(* IEC 61131-3 sources: daoli-st-library/DL_MathData (part 15) *)

(* ---- FC_DL_HexStringToLword.st ---- *)
(*==============================================================================
 * 组件名称 (Component)  : FC_DL_HexStringToLword
 * 所属子库 (Sublibrary) : DL_MathData
 * 归属目录 (Directory)  : C:\Library\DL_MathData
 * 当前版本 (Version)    : 1.0.0
 * 分类/来源标签         : 函数（FUNCTION）· 纯函数 · 十六进制串解析
 *                         iec-std-wrapper / string / bitstring
 * 兼容性   (Platform)   : CODESYS 3.5 / TwinCAT 3 / 汇川 InoProShop / 施耐德
 *                         Machine Expert；仅用 Standard.library 的 LEN / MID / FIND
 * 溯源声明 (Provenance) : IEC 61131-3 标准语义的道莅防御性实现——内部委托平台标准库语义，
 *                         外围统一错误码 / 钳位 / 双语注释，严禁重实现数学内核。
 * 功能一句话 (Summary)  : 大小写十六进制串解析为 LWORD，奇偶长度、非法字符、
 *                         超长溢出三闸齐备，与 FC_DL_BytesToHexString 互补成对。
 *
 * 功能描述 (Function)   : 一次锁存串长后按序过三闸：长度大于 16 即溢出闸、
 *                         奇数长度即对齐闸、逐字符经三张码表定位失败即非法闸；
 *                         合法路径每字符左移 4 位并入半字节，空串恒等返回零值。
 * 与既有件边界 (Boundary): 本件只解析裸十六进制串，不识别 0x 前缀、不下划线
 *                         分隔；超过 16 个有效位即溢出拒绝，绝不静默截高位。
 * 码位说明 (Codes)      : 信息 16#0002_3040 空输入恒等返回（值零、解析零位）
 *                         故障 16#0002_3041 奇数长度（半个字节无法对齐）
 *                         故障 16#0002_3042 非法字符（不在 0-9 A-F a-f）
 *                         故障 16#0002_3043 超长溢出（有效位大于 16）
 *                         段 16#02_3_40~43 首槽信息级、次槽起故障级。
 * 依赖说明 (Depends)    : 无 DL_ 内部依赖；仅 Standard.library 的 LEN / MID / FIND。
 * 红线自检 (Redline)    : 零全局依赖 ｜ 零 VAR_EXTERNAL ｜ 零 %I/%Q ｜ 纯 IEC 标准库
 *                         移位量 4 恒小于 64 位宽（归一达标）｜ 无除法面
 *                         全变量双语同行注释 ｜ 无定时器实例
 * 修订历史 (Revision)   : 2026-11-18  v1.0.0  首版入库（R32 · 批 1）
 *============================================================================*)

FUNCTION FC_DL_HexStringToLword : BOOL
VAR_INPUT
    sHex : STRING(255);                 // 源十六进制串 [ASCII]，有效位最多 16 / Source hex string, at most 16 digits
END_VAR
VAR_OUTPUT
    uValue  : LWORD;                    // 解析结果 [位串]，域外拒绝时保持零 / Parsed value, zero when refused
    nParsed : INT;                      // 成功解析的有效位数 [位] / Digits parsed on success
    uErrorId: UDINT;                    // 事件码，0 表示无事件 / Event code, zero means none
END_VAR
VAR
    cCh    : STRING(1);   // 当前字符 [字符] / Current character
    nLen   : INT;         // 锁存的源串长度 [字符]，R38 唯一锁存量 / Latched source length
    nVal   : INT;         // 当前半字节值 [值]，域 0 到 15 / Current nibble value, 0 to 15
    nPos   : INT;         // 码表定位结果 [索引]，1 起 / Table position, 1-based
    nI     : INT;         // 字符循环下标 [索引] / Character loop index
    uAcc   : LWORD;       // 累积值 [位串]，出口一次性赋给 uValue / Accumulator
    uCode  : UDINT;       // 码位暂存，出口单点写入 [码] / Code staging
END_VAR
VAR CONSTANT
    DL_HTL_MAXDIG : INT := 16;  // 有效位上限 [位]，LWORD 恰好 64 位 / Digit limit, LWORD is exactly 64 bits
    DL_HTL_ONE    : INT := 1;   // 单字符长度参数 [字符] / Single character length argument
END_VAR

(* 段 1｜输出预置与残留清除 / Pre-set and clear before any branch *)
FC_DL_HexStringToLword := FALSE;
uValue   := 16#0000_0000_0000_0000;
uAcc     := 16#0000_0000_0000_0000;
nParsed  := 0;
uErrorId := 16#0000_0000;
uCode    := 16#0000_0000;

(* 段 2｜LEN 一次锁存 / Latch the length once *)
nLen := LEN(sHex);
IF nLen < 0 THEN
    nLen := 0;                   // 防御：异常返回值钳到零 / Defensive clamp
END_IF

(* 段 3｜空串恒等：信息级告知后成功返回零值 / Empty string identity: inform and succeed *)
IF nLen = 0 THEN
    uErrorId := 16#0002_3040;    // 信息级：空输入恒等返回 / Info: empty input identity
    FC_DL_HexStringToLword := TRUE;
    RETURN;
END_IF

(* 段 4｜溢出闸：有效位超过 16 直接拒绝，绝不静默截高位 / Overflow gate: refuse, never truncate silently *)
IF nLen > DL_HTL_MAXDIG THEN
    uErrorId := 16#0002_3043;    // 故障级：超长溢出 / Fault: overflow by length
    RETURN;
END_IF

(* 段 5｜对齐闸：奇数长度意味着半个字节，解析结果无法定界 / Alignment gate: odd length leaves a half byte undefined *)
IF (nLen MOD 2) = 1 THEN
    uErrorId := 16#0002_3041;    // 故障级：奇数长度 / Fault: odd length
    RETURN;
END_IF

(* 段 6｜逐字符解析：三张码表定位，失败即非法闸 / Parse per character: three tables, failure is the legality gate *)
FOR nI := 1 TO nLen DO
    cCh := MID(sHex, DL_HTL_ONE, nI);                // 取当前字符 / Take the current character
    IF (cCh >= '0') AND (cCh <= '9') THEN
        nPos := FIND('0123456789', cCh);             // 数字表定位，域内恒 1 到 10 / Digit table, 1 to 10
        nVal := nPos - DL_HTL_ONE;                   // 值 0 到 9 / Value 0 to 9
    ELSIF (cCh >= 'A') AND (cCh <= 'F') THEN
        nPos := FIND('ABCDEF', cCh);                 // 大写表定位 / Uppercase table
        nVal := 10 + (nPos - DL_HTL_ONE);            // 值 10 到 15 / Value 10 to 15
    ELSIF (cCh >= 'a') AND (cCh <= 'f') THEN
        nPos := FIND('abcdef', cCh);                 // 小写表定位 / Lowercase table
        nVal := 10 + (nPos - DL_HTL_ONE);            // 值 10 到 15 / Value 10 to 15
    ELSE
        uErrorId := 16#0002_3042;                    // 故障级：非法字符 / Fault: illegal character
        RETURN;
    END_IF
    uAcc := SHL(uAcc, 4) OR INT_TO_LWORD(nVal);      // 左移 4 位并入半字节 / Shift four and OR the nibble
    nParsed := nParsed + DL_HTL_ONE;                 // 有效位计数 / Count the digit
END_FOR

(* 段 7｜出口装配：结果与码位单点写出 / Exit: single write for result and code *)
uValue := uAcc;
uErrorId := uCode;
FC_DL_HexStringToLword := TRUE;
END_FUNCTION

(* ---- FC_DL_HexToStr.st ---- *)
(*
  ==================================================================
  组件名 Component  : FC_DL_HexToStr
  分类   Category   : DL_MathData
  前缀   Naming     : FC_DL_ ｜ b/n/u/f/s/a 类型前缀制（R265）
  版本   Version    : 1.0.0
  功能   Purpose    : 字节串 → HEX 大写文本：每字节展开两位（高半字节
                      在前），输出上限 255 字符（2×127 字节 = 254 字符
                      + $00 终结符），超限按 R49 四步截断样板执行：先判
                      超限并置截断信息码与 bTrunc → 再钳长 → 再写入 →
                      最后显式写 $00 终结符。返回值 = 实际写入字符数
                      （名实双出口）。溯源：本件为「IEC 61131-3 标准语
                      义的道莅防御性实现」，内核委托标准库字符串函数
                      （MID/CONCAT/REPLACE/LEN），严禁重实现内核。
  来源   Source     : iec-std-wrapper（T0-6）：IEC 61131-3 标准语义的
                      道莅防御性实现，内核委托标准库字符串函数，零内核
                      重实现（T0-6 四步截断样板 R49）
  互引   Cross-ref  : FC_DL_StrToHex（同族逆变换件：HEX 文本 → 字节串，
                      二者成对使用需同参数约定：大写两位/字节、无分隔符）
  平台   Platform   : 纯 IEC 61131-3（标准库字符串函数 + SHR/MOD），三平台通用
  依赖   Depends    : 无 DL_ 内部依赖；标准字符串函数 MID/CONCAT/REPLACE/LEN
  设计偏差 Deviation: nLen 超出数组实际长度时按长度钳位接管（同族口径，
                      头注声明，不静默越界）；输出按 254 字符整字节截断
                      （255 上限内最大整字节边界，保证 $00 终结符可写）。
  红线   Redline    : R1 零全局/VAR_EXTERNAL/R2 零 %I/%Q/R3 纯 IEC 标准
                      R4 截断先判后钳（R49 四步）+ 终结符显式 + 下标界
                      闸/R5 全变量双语同行注释/R6 纯函数无状态机（CASE
                      不适用）/R7 无定时器与沿检测/R8 长度与查表界常量化
  错误码 Codes      : 01【信息级】超 255 字符上限截断（置 bTrunc，不置
                      bError，前缀字节完整保留）
                      02【失效级】nLen 超数组实际长度且钳位后为 0（无可
                      写字节），返回 0
  码位反证 Note     : 01/02 分立依据（R90）：01 在容量面（数据仍完整可
                      用，功能不受影响）、02 在输入面（无数据可转）可观
                      测；01 不置 bError 与 02 失效级双通道可区分。
  验收   Acceptance : V1 [0x0A,0xFF] → '0AFF' ｜ V2 [0x00] → '00' ｜
                      V3 128 字节 → 截断 127 字节 + bTrunc + 码 01 ｜
                      V4 nLen=0 → 空串（bValid）｜ V5 返回值 = LEN(sHexOut)
  变更   Revision   : 2026-11-22  v1.0.0  R67 首版（编码阶段批 2 序 5）
  ==================================================================
*)
FUNCTION FC_DL_HexToStr : UDINT
VAR_INPUT
    aBytes : ARRAY[*] OF BYTE;  // 输入字节串 [字节] / the input byte array
    nLen   : UDINT;             // 参与转换字节数 [字节]，超数组长度按长度钳位 / the byte count, clamped to the array length
END_VAR
VAR_OUTPUT
    sHexOut : STRING(255);      // HEX 大写文本（两位/字节，无分隔符）/ the hex uppercase text
    bTrunc  : BOOL;             // 截断标志（超 255 字符上限）[-] / the truncation flag
    bValid  : BOOL;             // 输出可用标志 [-] / the output usable flag
    nErrId  : UDINT;            // 错误码，0=正常，01/02 见头注 [码] / the error code [code]
END_VAR
VAR
    sHexTab : STRING := '0123456789ABCDEF'; // 半字节查表 [表] / the nibble lookup table
    sOut    : STRING(255);                  // 输出组装工作串 / the output assembly working string
    uUsed   : UDINT;                        // 钳位后实际字节数 [字节] / the used byte count after clamping
    uLenArr : UDINT;                        // aBytes 实际长度 [字节] / the actual array length
    i       : UDINT;                        // 字节遍历循环变量 / the byte loop index
    uB      : BYTE;                         // 当前字节工作寄存器 / the current byte register
    uHi     : BYTE;                         // 高半字节 [半字节] / the high nibble
    uLo     : BYTE;                         // 低半字节 [半字节] / the low nibble
    sCh     : STRING(1);                    // 当前查表字符 / the current looked up char
END_VAR
VAR CONSTANT
    H2S_CHARS_MAX : UDINT := UDINT#254;     // 输出字符上限（255 内整字节边界）[字符] / the output char ceiling
    H2S_BYTES_MAX : UDINT := UDINT#127;     // 对应字节数上限 [字节] / the matching byte ceiling
    H2S_ERR_NONE  : UDINT := 16#0000_0000;  // 无错误 [码] / no error [code]
    H2S_ERR_TRUNC : UDINT := 16#0000_0001;  // 码 01：超限截断（信息级）/ code 01, truncated, info level
    H2S_ERR_EMPTY : UDINT := 16#0000_0002;  // 码 02：无可写字节 / code 02, nothing to write
END_VAR

// 段 1｜输出预置 / segment 1, preset the outputs
sHexOut := '';                // 预置空串 / preset the empty string
bTrunc := FALSE;              // 预置未截断 / preset not truncated
bValid := FALSE;              // 预置不可用 / preset unusable
nErrId := H2S_ERR_NONE;       // 预置无错误 / preset no error
sOut := '';                   // 组装串清空 / clear the assembly string

// 段 2｜数组长度闸与钳位（结构性防御，头注偏差声明）/ segment 2, the array length clamp
IF UPPER_BOUND(aBytes, 1) >= 0 THEN
    uLenArr := DINT_TO_UDINT(1 + UPPER_BOUND(aBytes, 1) - LOWER_BOUND(aBytes, 1));  // 数组长度 / the array length
ELSE
    uLenArr := UDINT#0;
END_IF
uUsed := nLen;                // 先取原始字节数 / take the raw count
IF uUsed > uLenArr THEN
    uUsed := uLenArr;         // 超长钳位接管（头注偏差声明）/ clamp, documented deviation
END_IF

// 段 3｜R49 四步截断第 1 步：先判超限并置码置标志（赋值行前于钳位行）
//      segment 3, the truncation judged before clamping, the code precedes the clamp
IF 2 * uUsed > H2S_CHARS_MAX THEN
    bTrunc := TRUE;           // 截断标志 / the truncation flag
    nErrId := H2S_ERR_TRUNC;  // 信息级码（不置 bError）/ the info code, no fault flag
    uUsed := H2S_BYTES_MAX;   // 钳至整字节边界（254 字符）/ clamp to the whole byte boundary
END_IF

// 段 4｜零字节出口（码 02）：钳位后无可写 / segment 4, the zero byte exit
IF uUsed = UDINT#0 THEN
    nErrId := H2S_ERR_EMPTY;  // 无数据可转 / nothing to write
    sHexOut := '';            // 显式空串（含隐式终结符）/ the explicit empty string
    FC_DL_HexToStr := UDINT#0;  // 返回 0 字符（名实双出口）/ zero chars published
    RETURN;
END_IF

// 段 5｜逐字节展开（委托内核：SHR/MOD 取半字节 + MID 查表 + CONCAT 组装）
//      segment 5, the per byte expansion, the kernel delegated to the standard functions
FOR i := UDINT#0 TO uUsed - 1 DO
    uB  := aBytes[i];                              // 当前字节 / the current byte
    uHi := SHR(uB, 4);                             // 高半字节（移位量 4 < 位宽 8，R48 合规）/ the high nibble
    uLo := uB MOD 16;                              // 低半字节 / the low nibble
    sCh := MID(sHexTab, 1, BYTE_TO_DINT(uHi) + 1); // 高位查表（1 起位）/ the high lookup
    sOut := CONCAT(sOut, sCh);                     // 追加高位 / append the high char
    sCh := MID(sHexTab, 1, BYTE_TO_DINT(uLo) + 1); // 低位查表 / the low lookup
    sOut := CONCAT(sOut, sCh);                     // 追加低位 / append the low char
END_FOR

// 段 6｜R49 四步第 4 步：显式写 $00 终结符（REPLACE 标准函数，在 nChars+1 位）
//      segment 6, the explicit terminator write via the standard REPLACE
sHexOut := REPLACE(sOut, '$00', 1, 2 * uUsed + UDINT#1);  // 终结符落位（第 nChars+1 字符）/ the terminator placed

// 段 7｜出口映射（名实双出口：返回值 = 写入字符数）/ segment 7, the exit mapping
FC_DL_HexToStr := 2 * uUsed;  // 返回写入字符数 [字符] / the published char count
bValid := TRUE;               // 输出可用（截断仍可用，头注码 01 口径）/ usable, truncated still usable
END_FUNCTION

(* ---- FC_DL_HmsToTodChk.st ---- *)
(*
    FC_DL_HmsToTodChk —— 时 / 分 / 秒三分量合成 TOD（HMI 组态入口）
    ------------------------------------------------------------------
    组件名称  : FC_DL_HmsToTodChk
    分类      : DL_MathData / TimeOfDay
    前缀      : FC_DL_
    版本      : 1.0.0
    溯源      : IEC 61131-3 标准语义的道莅防御性实现（三分量组态合成 +
                域闸钳位口径）；TOD 合成内核**委托库内属主件
                FC_DL_DintMsToTod（DL_MathData，毫秒计数口径唯一属主）**，
                本件零内联 ms→TOD 转换（T0 委托纪律）；判据顺序与
                FC_DL_DurationFormat 域外钳位口径对齐（库内复用）；
                引脚名 / 码位 100% 自有；clean-room 声明 —— 零代码行复制。
    平台      : 纯 IEC 61131-3（UDINT 域闸 + 常量乘法 + 委托调用），
                CODESYS 3.5 / TwinCAT 3 / InoProShop / Machine Expert 通用
    作者      : 道莅代码库 · PLC编程专家（R72 构建轮 · 批 2 · 序号 6）
    ------------------------------------------------------------------
    功能说明  : HMI 三字段组态入口（时 / 分 / 秒各自独立输入）合成当日时刻
                TOD。真实工况：班次时刻 / 窗口时刻设定，与
                FB_DL_TimeWindowCheck / FB_DL_OccScheduleWindow 联用。
                判据链顺序：
                ① 分量非负闸：UDINT 天然非负，仅声明（无负值路径，闸空转）；
                ② 组合域闸（UDINT 域内先钳位后降位，防 UDINT→DINT 回绕）：
                   uHours > 23 → 钳 23；uMins > 59 → 钳 59；uSecs > 59 →
                   钳 59，**钳位照算 + 信息级**（与 FC_DL_DurationFormat 口径
                   对齐，不拒收——HMI 误输入尽量给出可用的最近合法时刻）；
                ③ 合成毫秒 nTotalMs = 时×3600000 + 分×60000 + 秒×1000：
                   上界推演 23×3600000 + 59×60000 + 59×1000 = 86399999
                   < 2^31 = 2147483648，钳位先行故乘法**无溢出面**（乘子全
                   常量，R382 常量除子 / 乘子级联口径）；
                ④ 委托属主件 FC_DL_DintMsToTod 合成 TOD（bClampSilently :=
                   TRUE——本件已钳到属主域 [0, 86399999] 内，属主钳位路径
                   结构性不可达），全 4 出参完整回执（R381 全回执纪律）；
                ⑤ 属主回执防御收口（回执不可用 → 故障级早退，结构性不可达）。
    错误码    : 16#0002_3909 分量越域（时 > 23 / 分 > 59 / 秒 > 59），已钳位
                            照算，bValid = TRUE —— 信息级，不置 bError（R45）
                16#0002_3910 属主件回执不可用（委托防御收口，结构性不可达）
                            —— 故障级
                加码反证句（R90）：3910 场景无法由 3909 + 正常返回观测——钳位
                路径 bValid = TRUE 且 TOD 有效，3910 是 bValid = FALSE 的
                不可用出口，输出组合不可互换观测，故立独立码。
    码位总账  : 16#0002_3909 用 ｜ 16#0002_3910 用
    状态机    : N/A —— 纯函数无状态，无 CASE 可写，非法状态不可能出现
    边界与披露: 一 无定时器 / 无沿检测实例 / 无数组下标 / 无除法（乘子常量
                   级联），周期安全规则 N/A；
                二 零全局变量、零 VAR_EXTERNAL、零物理地址；
                三 整数进位点（终审两式 #2）验收向量：「23:59:59 恰为上界」→
                   86399999 ms 正常出口不置码；「24:00:00 越界」→ 钳位
                   23:59:59 + 信息级 3909；
                四 域闸逐项点名（R272）：uHours / uMins / uSecs 三入参全部
                   纳入组合域闸，缺一即钳位静默失效；
                五 降位可表性：uHours ≤ 23 / uMins ≤ 59 / uSecs ≤ 59 已在
                   UDINT 域钳位后才 UDINT_TO_DINT，降位无回绕面（先钳后降
                   顺序写死，禁颠倒）；
                六 分工互引：FC_DL_TodToDintMs / FC_DL_DintMsToTod（毫秒计数
                   口径，后者为本件委托属主）、FC_DL_TimeToHmsString（TIME→
                   "hh:mm:ss" 文本）——本件为其组态侧反向语义，非文本变体；
                七 依赖声明：Standard.library（无内建函数依赖）+ 同库
                   FC_DL_DintMsToTod（只调用不修改）。
    验收向量  : V1 (8, 30, 0) → 08:30:00 正常出口；V2 (23, 59, 59) →
                86399999 ms 上界正常出口；V3 (24, 0, 0) → 钳位 23:59:59 +
                3909；V4 (0, 60, 0) → 钳位 00:59:00 + 3909；
                V5 (4294967295, 0, 0) → 钳位 23:00:00 + 3909（UDINT 域闸
                先行，降位无回绕向量）。
                算法已证（脚本）：未跑 ｜ 编译器已证（三平台）：未跑
    修订记录  : 2026-11-23 v1.0.0 首次入库（R72 构建轮 · 批 2 · 序号 6）
*)
FUNCTION FC_DL_HmsToTodChk : TOD
VAR_INPUT
    uHours : UDINT;                        (* 时分量，[时]，域 0~23，越域钳位照算 / the hours component, clamped outside *)
    uMins  : UDINT;                        (* 分分量，[分]，域 0~59，越域钳位照算 / the minutes component, clamped outside *)
    uSecs  : UDINT;                        (* 秒分量，[秒]，域 0~59，越域钳位照算 / the seconds component, clamped outside *)
END_VAR
VAR_OUTPUT
    bValid    : BOOL;                      (* 返回值（TOD）可用标志，故障级为 FALSE / the TOD usable flag *)
    bError    : BOOL;                      (* 故障标志，仅故障级码置位（R45 配对）/ the fault flag *)
    nInfoCode : UDINT;                     (* 信息 / 错误码，0 = 正常 / the info or error id *)
END_VAR
VAR CONSTANT
    DL_HMS_HMAX : UDINT := 23;             (* 时分量域上界 [时] / the hours domain upper bound *)
    DL_HMS_MMAX : UDINT := 59;             (* 分分量域上界 [分] / the minutes domain upper bound *)
    DL_HMS_SMAX : UDINT := 59;             (* 秒分量域上界 [秒] / the seconds domain upper bound *)
    DL_HMS_MSH  : DINT := 3600000;         (* 每小时毫秒数（常量乘子级联，R382）[ms] / the milliseconds per hour *)
    DL_HMS_MSM  : DINT := 60000;           (* 每分钟毫秒数 [ms] / the milliseconds per minute *)
    DL_HMS_MSS  : DINT := 1000;            (* 每秒毫秒数 [ms] / the milliseconds per second *)
END_VAR
VAR
    uHClamp : UDINT;                       (* 钳位后时分量 [时] / the clamped hours *)
    uMClamp : UDINT;                       (* 钳位后分分量 [分] / the clamped minutes *)
    uSClamp : UDINT;                       (* 钳位后秒分量 [秒] / the clamped seconds *)
    nH      : DINT;                        (* 降位时分量 [时] / the narrowed hours *)
    nM      : DINT;                        (* 降位分分量 [分] / the narrowed minutes *)
    nS      : DINT;                        (* 降位秒分量 [秒] / the narrowed seconds *)
    nTotalMs : DINT;                       (* 合成当日毫秒（上界 86399999 已证可表）[ms] / the composed day milliseconds *)
    _bMsErr : BOOL;                        (* 属主件故障回执 [标志] / the owner FC fault receipt *)
    _bMsVld : BOOL;                        (* 属主件输出可用回执（R381 全回执）[标志] / the owner FC usable receipt *)
    _bMsClmp: BOOL;                        (* 属主件钳位回执（结构性恒 FALSE，收下备用）[标志] / the owner FC clamp receipt *)
    _eMsCode: UDINT;                       (* 属主件码位回执 [码] / the owner FC code receipt *)
END_VAR

// 段 1｜返回值与状态预置（统一出口预置，R256）/ segment 1, preset the return and the status
FC_DL_HmsToTodChk := T#0S;                 // 故障缺省返回当日零点 / the fault default is midnight
bValid    := FALSE;                        // 预置不可用，过闸后置位 / preset unusable
bError    := FALSE;                        // 预置无故障 / preset no fault
nInfoCode := 0;                            // 预置无错 / preset no error
uHClamp := 0;                              // 钳位中间量清零 / clear the clamped hours
uMClamp := 0;                              // 钳位中间量清零 / clear the clamped minutes
uSClamp := 0;                              // 钳位中间量清零 / clear the clamped seconds
nH := 0;                                   // 降位中间量清零 / clear the narrowed hours
nM := 0;                                   // 降位中间量清零 / clear the narrowed minutes
nS := 0;                                   // 降位中间量清零 / clear the narrowed seconds
nTotalMs := 0;                             // 合成毫秒清零 / clear the composed milliseconds
_bMsErr := FALSE;                          // 属主回执清零 / clear the owner receipts
_bMsVld := FALSE;                          // 属主回执清零 / clear the owner receipts
_bMsClmp := FALSE;                         // 属主回执清零 / clear the owner receipts
_eMsCode := 0;                             // 属主码位清零 / clear the owner code

// 段 2｜分量非负闸（UDINT 天然非负，仅声明；无负值路径，闸空转）/ segment 2, the non negative declaration gate
// UDINT 域无负值路径，本闸为声明性空转（R272 全枚举中的口径声明行）。
// The UDINT domain has no negative path, this gate is a declarative no op.

// 段 3｜组合域闸：UDINT 域内先钳位后降位（防 UDINT→DINT 回绕，先钳后降顺序写死）/ segment 3, the combined domain gate with clamp before narrowing
IF uHours > DL_HMS_HMAX THEN               // 时越上界 / the hours over the bound
    uHClamp := DL_HMS_HMAX;                // 钳到 23 / clamp to 23
ELSE                                       // 时在域内 / the hours inside
    uHClamp := uHours;                     // 原值接管 / take the raw value
END_IF
IF uMins > DL_HMS_MMAX THEN                // 分越上界 / the minutes over the bound
    uMClamp := DL_HMS_MMAX;                // 钳到 59 / clamp to 59
ELSE                                       // 分在域内 / the minutes inside
    uMClamp := uMins;                      // 原值接管 / take the raw value
END_IF
IF uSecs > DL_HMS_SMAX THEN                // 秒越上界 / the seconds over the bound
    uSClamp := DL_HMS_SMAX;                // 钳到 59 / clamp to 59
ELSE                                       // 秒在域内 / the seconds inside
    uSClamp := uSecs;                      // 原值接管 / take the raw value
END_IF
IF (uHours > DL_HMS_HMAX) OR (uMins > DL_HMS_MMAX) OR (uSecs > DL_HMS_SMAX) THEN // 任一分量越域 / any component out of domain
    nInfoCode := 16#0002_3909;             // 信息级：钳位照算（DurationFormat 对齐口径）/ info level: clamped
    bError := FALSE;                       // 信息级不置故障（R45）/ info level never raises a fault
END_IF

// 段 4｜降位与毫秒合成（乘子全常量级联，上界 86399999 < 2^31 无溢出面）/ segment 4, narrowing and the millisecond composition
nH := UDINT_TO_DINT(uHClamp);              // 降位时分量（已证 <= 23）/ narrow the hours proven safe
nM := UDINT_TO_DINT(uMClamp);              // 降位分分量（已证 <= 59）/ narrow the minutes
nS := UDINT_TO_DINT(uSClamp);              // 降位秒分量（已证 <= 59）/ narrow the seconds
nTotalMs := (nH * DL_HMS_MSH) + (nM * DL_HMS_MSM) + (nS * DL_HMS_MSS); // 常量乘子合成 / the composition with constant multipliers

// 段 5｜委托属主件合成 TOD（返回值 TOD 直接承接；bClampSilently := TRUE，
//        属主钳位路径结构性不可达；全 4 出参完整回执，R381）/ segment 5, the delegated TOD composition
FC_DL_HmsToTodChk := FC_DL_DintMsToTod(nMsOfDay := nTotalMs, // 当日毫秒入参（已证在属主域内）/ the day milliseconds inside the owner domain
                                       bClampSilently := TRUE, // 钳位静默选向（本件已钳，属主钳位不可达）/ the silent clamp selector
                                       eErr => _eMsCode,       // 码位回执 / the code receipt
                                       bError => _bMsErr,      // 故障回执 / the fault receipt
                                       bValid => _bMsVld,      // 输出可用回执（R381 全回执）/ the usable receipt
                                       bClamped => _bMsClmp);  // 钳位回执 / the clamp receipt
IF _bMsErr OR (NOT _bMsVld) THEN           // 属主回执防御收口（结构性不可达）/ the owner receipt defensive guard
    nInfoCode := 16#0002_3910;             // 故障级：属主回执不可用 / fault level: the owner receipt unusable
    bError := TRUE;                        // R45 配对置故障标志 / paired with the fault flag
    bValid := FALSE;                       // 返回值不可用 / the return unusable
    FC_DL_HmsToTodChk := T#0S;             // 确定值零点出口 / a deterministic midnight outlet
    RETURN;                                // 结构早退 / structural exit
END_IF

// 段 6｜正常出口 / segment 6, the normal outlet
bValid := TRUE;                            // 结果可用 / the result usable
END_FUNCTION

(* ---- FC_DL_HoneCrosshatchAngleCalc.st ---- *)
(*
  DL Factory R88 | FC_DL_HoneCrosshatchAngleCalc
  功能：由往复速度与旋转线速度算珩磨网纹夹角 θ=2·atan(vr/vt)，按 20°~60° 判带宽
  开源溯源：无（clean-room 自研，依据公开工艺公式 珩磨网纹角式 θ=2·atan(vr/vt)，许可证=MIT，借鉴点=公式结构）
  规则：R1-R16 全遵守；R88 简单件标量形（纯标量入参出参，无循环体、无方法、无属性、无数组）
*)
FUNCTION FC_DL_HoneCrosshatchAngleCalc : REAL
VAR_INPUT
    fRecipSpeedMPerMin : REAL := 15.0; // 珩磨头往复速度 vr [m/min] / reciprocating speed [m/min]
    fRotSpeedMPerMin : REAL := 45.0; // 工件旋转线速度 vt（按孔径处分度线速度折算） [m/min] / rotational surface speed [m/min]
    fBandMinDeg : REAL := 20.0; // 网纹角允许下限（工艺带宽） [°] / lower crosshatch band [deg]
    fBandMaxDeg : REAL := 60.0; // 网纹角允许上限（工艺带宽） [°] / upper crosshatch band [deg]
END_VAR
VAR_OUTPUT
    fAngleDeg : REAL; // 网纹夹角 θ [°] / crosshatch included angle [deg]
    xInBand : BOOL; // TRUE=网纹角落在允许带宽内 [-] / TRUE when the angle is inside the band [-]
END_VAR
VAR
    fRatio : REAL; // 速度比 vr/vt（正切值） [-] / speed ratio, the tangent value [-]
    fAngleRad : REAL; // 半网纹角 atan(vr/vt) [rad] / half crosshatch angle [rad]
    fDenom : REAL; // 分母 vt（除零判据） [m/min] / denominator before the division [m/min]
END_VAR

// 段 1｜出口预置
FC_DL_HoneCrosshatchAngleCalc := -1.0; // 哨兵返回 -1（无效） [-] / sentinel return -1, invalid [-]
fAngleDeg := 0.0; // 网纹角预置零 [°] / angle preset zero [deg]
xInBand := FALSE; // 带宽位预置 FALSE [-] / band flag preset false [-]
fRatio := 0.0; // 速度比预置零 [-] / ratio preset zero [-]
fAngleRad := 0.0; // 半角预置零 [rad] / half angle preset zero [rad]
fDenom := 0.0; // 分母预置零 [m/min] / denominator preset zero [m/min]

// 段 2｜非有限拦截 + 域闸
IF NOT (fRecipSpeedMPerMin > -1.0E30 AND fRecipSpeedMPerMin < 1.0E30) OR NOT (fRotSpeedMPerMin > -1.0E30 AND fRotSpeedMPerMin < 1.0E30) THEN
    RETURN; // 两速度任一非有限即拒算 [-] / any non finite speed rejected [-]
END_IF
IF NOT (fBandMinDeg > -1.0E30 AND fBandMinDeg < 1.0E30) OR NOT (fBandMaxDeg > -1.0E30 AND fBandMaxDeg < 1.0E30) THEN
    RETURN; // 带宽上下限任一非有限则判据静默失效，故先拦 [-] / band limits must be finite or the check fades [-]
END_IF
IF fRecipSpeedMPerMin < 0.0 OR fRotSpeedMPerMin <= 0.0 THEN
    RETURN; // 往复速度非负闸 + 旋转速度正域闸（分母不得为零） [m/min] / non negative vr and positive vt [m/min]
END_IF
IF fBandMinDeg <= 0.0 OR fBandMaxDeg <= fBandMinDeg THEN
    RETURN; // 带宽自洽闸：下限须为正、上限须严格大于下限 [°] / band consistency gate [deg]
END_IF

// 段 3｜计算
fDenom := fRotSpeedMPerMin; // 取旋转线速度作除数 [m/min] / take the rotational speed as divisor [m/min]
IF fDenom < 1.0E-9 THEN
    RETURN; // 除法前分母闸：vt 必须大于 1E-9 才可作除数 [m/min] / denominator gate before the division [m/min]
END_IF
fRatio := fRecipSpeedMPerMin / fDenom; // (m/min) ÷ (m/min) = 无量纲 [-] / dimensionless ratio [-]
fAngleRad := ATAN(fRatio); // 无量纲 → 弧度，半网纹角 [rad] / half angle in radians [rad]
fAngleDeg := 2.0 * fAngleRad * 57.2957795; // 2 × rad × (180/π) = 度，换算常数 57.2957795 [°] / radians to degrees [deg]

// 段 4｜判定与饱和
IF NOT (fAngleDeg > -1.0E30 AND fAngleDeg < 1.0E30) THEN
    RETURN; // 结果非有限再拦一次 [-] / re-check the result for finiteness [-]
END_IF
xInBand := (fAngleDeg >= fBandMinDeg) AND (fAngleDeg <= fBandMaxDeg); // 双侧闭区间直比 [°] / closed two sided band compare [deg]

// 段 5｜出口自检
IF fAngleDeg <= 0.0 THEN
    RETURN; // 出口自检：网纹角须为正（零值说明往复速度为零） [°] / angle must be positive [deg]
END_IF
FC_DL_HoneCrosshatchAngleCalc := fAngleDeg; // 返回网纹夹角 θ [°] / return the crosshatch angle [deg]
END_FUNCTION

(* ---- FC_DL_Hypot3D.st ---- *)
(*
  ==================================================================
  组件名 Component  : FC_DL_Hypot3D
  分类   Category   : DL_MathData
  前缀   Naming     : FC_DL_ ｜ b/n/u/f/t/e/st 类型前缀制（R265）
  复杂度 Complexity  : 低
  版本   Version    : 1.0.0
  功能   Purpose    : 三维矢量模长 √(x²+y²+z²)，中途缩放防 x² 溢出。
  来源   Source     : self-std（公开数学语义自研包装）
  平台   Platform   : 纯 IEC 61131-3（SQRT / ABS / 四则运算），三平台通用
  分工声明 Split     : 与 FC_DL_Hypot（二维属主，若在册）互引——本件只做三维；
                      T0 防御性包装：内核即 SQRT 一次委托，不重实现数学内核。
  作者   Author     : 道莅代码库 · PLC 编程专家（R61）
  归属 Ownership     : 本件无 TYPE 声明；引用件类型全部 IEC 标准原生。
  ------------------------------------------------------------------
  边界 Boundary     :
                      一 非有限闸逐个点名三个浮点入参（R272 全量枚举：fX / fY /
                         fZ 三个各判 NaN 自反 + Inf 差值自减），命中即拒绝出值；
                      二 溢出防护：先取三轴绝对值最大者 fMax 缩放，归一化分量
                         |fXn| ≤ 1，平方和 ≤ 3 结构性不溢出，再乘回 fMax；
                      三 全零矢量：fMax = 0 时直接返回 0（禁除零，除子已证 > 0）；
                      四 结果复检兜底同拍置 eErr + bError + bValid 三件套（R258）；
                      五 无状态纯函数：局部量段 1 显式预置（R254）。
  错误码   Codes    :
    16#0001_0631【故障级】入参含非有限值（fX / fY / fZ 逐个点名），拒绝出值
    16#0001_0632【故障级】结果非有限（复检兜底，结构性不可达仍保留）
  验收   Acceptance :
    算法已证（脚本）：未跑 ｜ 编译器已证（三平台）：未跑
    V1 (3,4,0) → 5.0；V2 (1E200,1E200,1E200) → 缩放后 ≈1.7320508E200 不溢出
    V3 fX=NaN → 码 0631、bValid=FALSE、返回 0
  修订记录 Revision  :
    2026-11-21  v1.0.0  R61 首版（批 1 · 序号 3）
  ==================================================================
*)
FUNCTION FC_DL_Hypot3D : LREAL
VAR_INPUT
    fX : LREAL; // X 分量 [用户单位] / the X component
    fY : LREAL; // Y 分量 [用户单位] / the Y component
    fZ : LREAL; // Z 分量 [用户单位] / the Z component
END_VAR
VAR_OUTPUT
    bValid : BOOL;  // 结果可用标志 [-] / the result usable flag
    eErr   : UDINT; // 错误码，0 = 正常 / the error code, zero is ok
    bError : BOOL;  // 错误标志，故障级码置位（R45 配对）/ the error flag
END_VAR
VAR
    fMax : LREAL; // 三轴绝对值最大者 [用户单位] / the largest absolute component
    fXn  : LREAL; // 归一化 X 分量 [-] / the normalised X component
    fYn  : LREAL; // 归一化 Y 分量 [-] / the normalised Y component
    fZn  : LREAL; // 归一化 Z 分量 [-] / the normalised Z component
END_VAR

// 段 1｜返回值与错误状态预置安全值（四段式第一段，R45）+ 局部量显式预置（R254）/ segment 1, the preset
FC_DL_Hypot3D := 0.0; // 返回值预置安全值零 / preset the return zero
bValid := FALSE; // 有效标志预置假 / preset the validity false
eErr := 16#0000_0000; // 错误码预置正常 / preset the code to ok
bError := FALSE; // 错误标志预置假 / preset the error flag false
fMax := 0.0; // 最大分量预置零 / preset the max zero
fXn := 0.0; // 归一化 X 预置零 / preset the normalised X zero
fYn := 0.0; // 归一化 Y 预置零 / preset the normalised Y zero
fZn := 0.0; // 归一化 Z 预置零 / preset the normalised Z zero

// 段 2｜非有限闸：三个入参逐个点名（R272 全量，边界一）/ segment 2, the finiteness gate naming every input
IF (fX <> fX) OR ((fX - fX) <> (fX - fX))
OR (fY <> fY) OR ((fY - fY) <> (fY - fY))
OR (fZ <> fZ) OR ((fZ - fZ) <> (fZ - fZ)) THEN // 任一分量非有限 / any component is not finite
    eErr := 16#0001_0631; // 故障级：入参含非有限值 / fault grade, a non finite input
    bError := TRUE; // 置错误标志（R45 配对）/ raise the error flag
    bValid := FALSE; // 结果不可用 / the result void
    RETURN; // 早退 / early return
END_IF

// 段 3｜缩放防溢出：先取最大绝对值（边界二）/ segment 3, the scaling against the overflow
fMax := ABS(fX); // 以 X 绝对值起步 / start from the absolute X
IF ABS(fY) > fMax THEN // Y 更大 / the Y is larger
    fMax := ABS(fY); // 接管最大值 / take over the max
END_IF
IF ABS(fZ) > fMax THEN // Z 更大 / the Z is larger
    fMax := ABS(fZ); // 接管最大值 / take over the max
END_IF
IF fMax = 0.0 THEN // 全零矢量（整数零精确比较，非浮点容差场景）/ the all zero vector with an exact integer zero compare
    FC_DL_Hypot3D := 0.0; // 模长为零 / the length is zero
    bValid := TRUE; // 结果可用 / the result is usable
    FC_DL_Hypot3D := 0.0; // 返回零 / return zero
ELSE // 非零矢量：归一化后开方再乘回 / the nonzero vector
    fXn := fX / fMax; // 归一化 X（除子 fMax 已证 > 0）/ the normalised X with a proven divisor
    fYn := fY / fMax; // 归一化 Y / the normalised Y
    fZn := fZ / fMax; // 归一化 Z / the normalised Z
    FC_DL_Hypot3D := fMax * SQRT(fXn * fXn + fYn * fYn + fZn * fZn); // 模长（平方和 ≤ 3 结构性不溢出）/ the length, the sum of squares bounded by three
END_IF

// 段 4｜结果复检兜底（非有限同拍三件套，边界四）/ segment 4, the result recheck
IF (FC_DL_Hypot3D <> FC_DL_Hypot3D)
OR ((FC_DL_Hypot3D - FC_DL_Hypot3D) <> (FC_DL_Hypot3D - FC_DL_Hypot3D)) THEN // 结果非有限 / the result is not finite
    FC_DL_Hypot3D := 0.0; // 兜底安全值 / the bottom line safe value
    eErr := 16#0001_0632; // 故障级：结果非有限 / fault grade, the non finite result
    bError := TRUE; // 置错误标志（R45 配对）/ raise the error flag
    bValid := FALSE; // 结果不可用 / the result void
ELSE // 结果有限 / a finite result
    bValid := TRUE; // 结果可用 / the result is usable
END_IF
END_FUNCTION

(* ---- FC_DL_HypotChk.st ---- *)
(*==============================================================================
 * 名称 : FC_DL_HypotChk —— 2D 斜边（max/min 比值缩放法防中间量溢出）
 * 分类 / 前缀 / 版本 : DL_MathData / FC_DL_ / 1.0.0
 * 溯源 : 开源语义参考（OSCAT/AixOCAT 族，MIT）或 clean-room IEC 实现，未复制源码
 * 平台 : 纯 IEC 61131-3
 * 功能说明 : 返回 sqrt(x^2 + y^2)，采用缩放算法：取 a=max(|x|,|y|)、
 *            b=min(|x|,|y|)，结果 = a*sqrt(1+(b/a)^2)。中间量 (b/a)^2 <= 1
 *            有界，杜绝直接 x^2+y^2 在大输入（如 1.0E200）下的中间溢出。
 *            边界处理：任一输入非有限（NaN/±Inf）置 eErr 返回 0.0；两输入
 *            全 0 时返回 0.0（合法结果，bValid 保持 TRUE）。
 * 错误码 : 16#0001_1B10 = 输入非有限（NaN/±Inf）
 *          eErr=0 且 bValid=TRUE 表示返回值可用
 * 状态机 : R6 标注 N/A（纯函数无顺序状态，以本节替代 ELSE 兜底）
 * 红线 : R1/R2/R3 ✓ 零全局/零IO/纯IEC ｜ R4 ✓ 非有限拦截/缩放防溢出/除零防护（a=0 特判）｜ R10 ✓ 标准转换 ｜ R11 ✓ 分号收尾 ｜ R15 ✓ 无保留字撞名
 * 修订记录 : 2026-11-23 v1.0.0 首次入库（R76）
 *============================================================================*)
FUNCTION FC_DL_HypotChk : LREAL
VAR_INPUT
    fX : LREAL;    // 直角边 X [工程单位] / leg X
    fY : LREAL;    // 直角边 Y [工程单位] / leg Y
END_VAR
VAR_OUTPUT
    eErr   : UDINT;    // 故障码，0=正常，1B10=输入非有限 / error code
    bError : BOOL;     // TRUE=本件发生故障 / TRUE when fault occurred
    bValid : BOOL;     // TRUE=返回值可用 / TRUE when return value is usable
END_VAR
VAR
    _fA : LREAL;       // 较大边（缩放基准）[工程单位] / larger leg as scale base
    _fB : LREAL;       // 较小边 [工程单位] / smaller leg
    _fR : LREAL;       // b/a 比值 [无量纲] / ratio b/a, bounded by 1
END_VAR

FC_DL_HypotChk := 0.0;                       // 返回值预设 0.0 / preset return to zero
eErr   := 16#0000_0000;                      // 故障码清零 / clear error code
bError := FALSE;                             // 故障标志清零 / clear error flag
bValid := TRUE;                              // 预设输出可用 / preset valid flag

IF (fX <> fX) OR ((fX - fX) <> (fX - fX))    // fX 非有限 / fX is NaN or infinite
   OR (fY <> fY) OR ((fY - fY) <> (fY - fY)) THEN    // fY 非有限 / fY is NaN or infinite
    eErr   := 16#0001_1B10;                  // 置非有限故障码 / set non-finite code
    bError := TRUE;                          // 置故障标志 / set error flag
    bValid := FALSE;                         // 返回值不可用 / return not usable
    RETURN;                                  // 返回 0.0 / return zero
END_IF

IF ABS(fX) >= ABS(fY) THEN                   // 按绝对值定大小序 / order by absolute value
    _fA := ABS(fX);                          // 大边 = |fX| / larger leg
    _fB := ABS(fY);                          // 小边 = |fY| / smaller leg
ELSE                                         // 反之 / otherwise
    _fA := ABS(fY);                          // 大边 = |fY| / larger leg
    _fB := ABS(fX);                          // 小边 = |fX| / smaller leg
END_IF

IF _fA = 0.0 THEN                            // 两边全 0：斜边 0（合法）/ both zero: hypot 0
    FC_DL_HypotChk := 0.0;                   // 返回 0.0 / return zero
    RETURN;                                  // 提前收口（防下步除零）/ early exit guards division
END_IF

_fR := _fB / _fA;                            // 比值 <=1，有界无溢出 / ratio bounded by one
FC_DL_HypotChk := _fA * SQRT(1.0 + _fR * _fR);    // 缩放法合成斜边 / scaled hypot

END_FUNCTION

(* ---- FC_DL_Hysteresis.st ---- *)
(*==============================================================================
 * 组件名称 (Component)  : FC_DL_Hysteresis
 * 所属子库 (Sublibrary) : DL_MathData
 * 当前版本 (Version)    : 1.0.0
 * 兼容性   (Platform)   : CODESYS 3.5 / TwinCAT 3 / 汇川 InoProShop / Machine Expert
 *                         仅依赖 Standard.library（ABS），全 REAL 运算
 * 功能描述 (Function)   : 施密特迟滞比较器（双阈值）。输入高于上阈值置 TRUE、
 *                         低于下阈值置 FALSE、落入回差带内保持原态。
 *                         用于液位、温度、压力等模拟量驱动的泵 / 加热器 / 报警器启停，
 *                         消除单阈值在设定点附近反复跨越导致的高频动作。
 *
 * 【接口设计决策 / Interface decision】
 *   迟滞的输出依赖上一周期输出，本质是有状态运算。本组件保持 FC_ 形态（不用 FB），
 *   状态经 VAR_IN_OUT bState 交还调用方持有：调用方声明持久变量 bHystState : BOOL;
 *   并每个扫描周期传入同一变量。好处是无实例内存、可直接放进 IF 表达式；
 *   代价是调用方必须遵守"同一变量回传"纪律。
 *
 * 【有状态纪律警告 / State retention warning（边界 B7）】
 *   VAR_IN_OUT 传入的必须是持久变量（实例成员、静态变量或 RETAIN 变量）。
 *   禁止传表达式、常量或临时变量，否则每周期状态被重置，退化为纯比较器：
 *     ✗ 错误示例：bPump := FC_DL_Hysteresis(fIn := fLevel, fThreshold := 60.0,
 *                                          fHysteresis := 2.0, bState := FALSE);
 *     ✓ 正确示例：bPump := FC_DL_Hysteresis(fIn := fLevel, fThreshold := 60.0,
 *                                          fHysteresis := 2.0, bState := bLevelHystState);
 *
 * 【初值行为 / Initial state behavior（边界 B5）】
 *   bState 上电初值 FALSE，若输入一开始就落在回差带内，输出保持 FALSE 不误动作
 *   （保守方向对泵与加热器均为安全侧）。若需"首次强制同步"，可先用一个低于下阈值的
 *   假值空跑一个周期，使状态与真实工况对齐。
 * 开源溯源 (Origin)     : 原创实现。施密特触发器为公开经典电路模型，本处为其离散化。
 * 依赖     (Depends)    : 无 DL_ 内部依赖
 * 红线自检 (Redline)    : R1 ✓ 零全局变量表与外部变量引用 ｜ R2 ✓ 零物理 IO 地址直写
 *                         R3 ✓ 纯 IEC 61131-3 ｜ R4 ✓ 负宽容错 + 回差上限 + 零回差告警 + 容差判零
 *                         R5 ✓ 全变量中英双语同行注释 + 有状态纪律警告 ｜ R6 N/A（用状态位非状态机）
 *                         R7 N/A（无定时器/边沿实例）
 * 修订历史 (Revision)   :
 *   2026-11-14  v1.0.0  首版入库（Phase 1 冷启动 · Level 0 批次）
 *============================================================================*)
FUNCTION FC_DL_Hysteresis : BOOL
VAR_INPUT
    fIn         : REAL;           // 输入值 [EU] / Input value [EU]
    fThreshold  : REAL;           // 设定点，回差带中心 [EU] / Setpoint, center of the hysteresis band [EU]
    fHysteresis : REAL := 0.0;    // 回差总宽度 [EU]，负值取绝对值 / Total hysteresis width [EU], negative taken as absolute
END_VAR
VAR_IN_OUT
    bState      : BOOL;           // 迟滞状态，调用方持有并每周期回传同一变量 / Hysteresis state, retained by the caller
END_VAR
VAR_OUTPUT
    fUpperTrip  : REAL;           // 实际上阈值 = fThreshold + 半回差 [EU] / Effective upper trip [EU]
    fLowerTrip  : REAL;           // 实际下阈值 = fThreshold - 半回差 [EU] / Effective lower trip [EU]
    uErrorId    : UDINT;          // 故障码，0 = 无故障 / Error code, 0 = no error
END_VAR
VAR
    fHalfBand      : REAL;        // 半回差带宽 [EU] / Half hysteresis band [EU]
    fThresholdAbs  : REAL;        // 设定点绝对值 [EU] / Absolute value of the setpoint [EU]
    fMaxBand       : REAL;        // 半回差允许上限 [EU] / Upper limit of the half band [EU]
END_VAR
VAR CONSTANT
    DL_FLOAT_EPS      : REAL := 1.0E-6;  // 浮点判零容差 / Float zero tolerance
    DL_HYST_MAX_RATIO : REAL := 0.5;     // 回差不超过设定点绝对值的 50%，防误填 / Max hysteresis ratio
END_VAR

(*------------------------------------------------------------------------------
 * 段 1｜默认保持原态：本函数在回差带内"什么都不做"，这是迟滞的定义
 *      Default hold: inside the band nothing is written, which is the definition
 *-----------------------------------------------------------------------------*)
FC_DL_Hysteresis := bState;
uErrorId         := 16#0000_0000;
fHalfBand        := 0.0;
fMaxBand         := 0.0;

(*------------------------------------------------------------------------------
 * 段 2｜回差负值容错（边界 B1）：取绝对值继续运行，仅告警
 *      Negative hysteresis tolerance: absolute value plus a warning only
 *-----------------------------------------------------------------------------*)
fHalfBand := ABS(fHysteresis) * 0.5;

IF fHysteresis < 0.0 THEN
    uErrorId := 16#0001_0003;
END_IF

(*------------------------------------------------------------------------------
 * 段 3｜回差上限保护（边界 B2）：按设定点绝对值的比例限幅
 *      Hysteresis upper limit: ratio based on the absolute setpoint value
 *      设定点本身接近 0 时相对上限退化（任何比例乘 0 都是 0），此时跳过比例限幅，
 *      否则回差会被压成 0、迟滞功能被静默取消
 *      限幅目的：防止参数误填导致阈值跑到物理量程之外、设备永不动作
 *-----------------------------------------------------------------------------*)
fThresholdAbs := ABS(fThreshold);

IF fThresholdAbs > DL_FLOAT_EPS THEN
    fMaxBand := fThresholdAbs * DL_HYST_MAX_RATIO;

    IF fHalfBand > fMaxBand THEN
        fHalfBand := fMaxBand;
        uErrorId  := 16#0001_0003;
    END_IF
END_IF

(*------------------------------------------------------------------------------
 * 段 4｜双阈值计算：上下阈值对称分布于设定点两侧
 *      Dual threshold computation, symmetric around the setpoint
 *-----------------------------------------------------------------------------*)
fUpperTrip := fThreshold + fHalfBand;
fLowerTrip := fThreshold - fHalfBand;

(*------------------------------------------------------------------------------
 * 段 5｜迟滞判定（边界 B3/B4）：置位用严格大于、复位用严格小于
 *      Hysteresis decision: strict greater for set, strict less for reset
 *      等于阈值时保持原态——写成 >= / <= 会让回差带退化，边界抖动立刻回来
 *      零回差时退化为普通比较器，允许运行但必须告警（组态缺陷而非运行故障）
 *-----------------------------------------------------------------------------*)
IF fHalfBand <= DL_FLOAT_EPS THEN
    (* 零回差：阈值重合，按严格不等式做单阈值比较，并置告警 *)
    (* Zero hysteresis: thresholds coincide, single-threshold comparison with a warning *)
    uErrorId := 16#0001_0003;

    IF fIn > fThreshold THEN
        bState := TRUE;
    ELSIF fIn < fThreshold THEN
        bState := FALSE;
    END_IF
ELSE
    IF fIn > fUpperTrip THEN
        bState := TRUE;
    ELSIF fIn < fLowerTrip THEN
        bState := FALSE;
    END_IF
END_IF

(*------------------------------------------------------------------------------
 * 段 6｜结果回写：同时返回更新后的状态，便于调用方在一次扫描内使用
 *      Result write-back: also return the refreshed state for same-scan use
 *-----------------------------------------------------------------------------*)
FC_DL_Hysteresis := bState;
END_FUNCTION

(* ---- FC_DL_IndexClampEx.st ---- *)
(*
    FC_DL_IndexClampEx —— 数组下标钳位原子（DINT 域）
    ------------------------------------------------------------------
    分类      : DL_MathData / Clamp
    前缀      : FC_DL_
    版本      : 1.0.0
    溯源      : IEC 61131-3 标准语义的道莅防御性实现
                （内部委托比较与选择语义，外围统一错误码/钳位/双语文档；
                  未复制任何闭源厂商源码，参考实现仅限 MIT/Apache 许可）
    平台      : 纯 IEC 61131-3，CODESYS / TwinCAT / InoProShop 通用
    作者      : 道莅代码库 · PLC编程专家（R40）
    ------------------------------------------------------------------
    功能说明  : 数组下标钳位原子：将 nIdx 钳制到 [nLower, nUpper] 边界内并作为
                返回值输出，供全部数组访问前的防御性下标整备复用；
                越界按边界钳位：nIdx < nLower 钳至下界，置信息级 16#0001_049C；
                nIdx > nUpper 钳至上界，置信息级 16#0001_049D；
                上下界倒置（nLower > nUpper）判为故障级 16#0001_03DA，返回下界值
                且 bValid=FALSE（倒置边界意味着调用方组态错误，钳位结果无确定
                语义，拒绝输出并保持返回值落在下界侧防御值）；
                信息级码属正常防御：bError=FALSE、bValid=TRUE，输出钳位后防御值。
    错误码    : 16#0001_03DA 上下界倒置（nLower > nUpper）——故障级，返回下界值，bValid=FALSE
                16#0001_049C 下标低于下界，已钳至下界——信息级，正常防御
                16#0001_049D 下标高于上界，已钳至上界——信息级，正常防御
                （R90 反证句：下越界与上越界两场景均无法由返回值观测——钳位后输出
                  为合法边界值且 bValid=TRUE 与域内直通组合相同，若不占码则现场无法
                  还原越界方向，故两侧各占一码；倒置场景由 bValid=FALSE 加故障码
                  组合与信息级钳位区分，且与两个越界码的「方向语义」不同，故独立占码）
    状态机    : R6 标注 N/A —— 本组件为纯函数无顺序状态机，无 CASE 可写，
                非法状态不可能出现，故以本节说明替代 ELSE 兜底
    修订记录  : 2026-11-19 v1.0.0 首次入库（R40 · 批 4 · T0 快车道）
*)
FUNCTION FC_DL_IndexClampEx : DINT
VAR_INPUT
    nIdx    : DINT; // 待钳位下标 [索引] ｜ index to clamp
    nLower  : DINT; // 边界下界 [索引]，大于上界时判故障拒绝 ｜ lower bound, a fault is raised when greater than the upper bound
    nUpper  : DINT; // 边界上界 [索引]，小于下界时判故障拒绝 ｜ upper bound, a fault is raised when less than the lower bound
END_VAR
VAR_OUTPUT
    eErr   : UDINT; // 错误码，0=正常，16#0001_04XX=信息级，16#0001_03XX=故障级 ｜ error id, 0=ok, 16#0001_04XX=info, 16#0001_03XX=fault
    bError : BOOL;  // 是否出错，eErr 落故障级时为 TRUE ｜ fault flag, TRUE when eErr is fault level
    bValid : BOOL;  // 输出是否有效可用 ｜ output valid flag
END_VAR

// 段 1｜返回值与错误状态预置 ｜ segment 1, preset return value and error status
FC_DL_IndexClampEx := 0; // 故障缺省返回 0 [索引] ｜ fault default returns 0
eErr   := 0;     // 预置无错误 ｜ preset no error
bError := FALSE; // 预置无故障 ｜ preset no fault
bValid := FALSE; // 预置无效，通过防御闸后置位 ｜ preset invalid, set TRUE after guard passes

// 段 2｜上下界倒置防御闸（早退） ｜ segment 2, bound-inversion guard (early return)
IF nLower > nUpper THEN
    FC_DL_IndexClampEx := nLower; // 故障级返回下界侧防御值 [索引] ｜ fault level returns the lower-bound defensive value
    eErr   := 16#0001_03DA;       // 上下界倒置故障码 ｜ bound-inversion fault id
    bError := TRUE;               // 置故障标志（R45 配对）｜ raise the fault flag (R45 pairing)
    bValid := FALSE;              // 输出无效 ｜ output invalid
    RETURN;                       // 早退，不做钳位推断 ｜ early return, no clamping inference
END_IF

// 段 3｜双侧钳位主体（末段） ｜ segment 3, double-side clamp body (final)
IF nIdx < nLower THEN
    FC_DL_IndexClampEx := nLower; // 低于下界钳至下界 [索引] ｜ under the lower bound, clamp to it
    eErr := 16#0001_049C;         // 信息级：下越界已钳位 ｜ info level: under-range clamped
ELSIF nIdx > nUpper THEN
    FC_DL_IndexClampEx := nUpper; // 高于上界钳至上界 [索引] ｜ over the upper bound, clamp to it
    eErr := 16#0001_049D;         // 信息级：上越界已钳位 ｜ info level: over-range clamped
ELSE
    FC_DL_IndexClampEx := nIdx;   // 域内下标直通 [索引] ｜ in-domain index pass-through
END_IF
bError := FALSE; // 信息级钳位不置故障，故障分支已提前返回 ｜ info-level clamp never raises fault, fault branch has returned
bValid := TRUE;  // 域内或钳位输出均有效可用 ｜ in-domain or clamped output is valid
END_FUNCTION

(* ---- FC_DL_IntDigitCountUdint.st ---- *)
(*==============================================================================
 * 组件名称 : FC_DL_IntDigitCountUdint ｜ 子库 : DL_MathData ｜ v1.0.0 ｜ 2026-11-24
 * 平台     : CODESYS 3.5 / TwinCAT 3 / InoProShop / Machine Expert（纯 IEC，无厂商库）
 * 功能简介 : 无符号整数的十进制位数（0 计 1 位）。循环整除 10 计数，纯整数实现，
 *            不使用字符串转换 —— 各平台 INT_TO_STRING 的前导空格/补零口径互不相同。
 * 契约     : 返回 1~10（UDINT 十进制最大 10 位）；nVal = 0 返回 1。
 * 依赖     : 无 DL_ 内部依赖（R16 自足实现），无标准库函数调用
 * 错误码   : R297 零码位范式：eErr 恒 0，仅以 bError / bValid 表达（本件结构性不置 bError）
 * 红线自检 : R1 零全局 R2 零%I/%Q R3 纯IEC R4 除数为常量 10、循环上界固定
 *            R5 双语注释 R6 N/A（无状态机）R7 N/A（无定时器/沿实例）
 *            R10 无类型转换 R11 全声明行分号 R15 标识符零保留字冲突 R18 N/A（无 bReset）
 * 修订历史 : 2026-11-24 R79-A 首版（整数数论族 4/8）
 *============================================================================*)
FUNCTION FC_DL_IntDigitCountUdint : UDINT
VAR_INPUT
    nVal        : UDINT;    // 待测位数的整数，全域 0~16#FFFF_FFFF [无量纲] / value whose decimal width is requested
END_VAR
VAR_OUTPUT
    eErr        : UDINT;    // 错误码，零码位范式恒 0 / error id, always zero under the zero-code rule
    bError      : BOOL;     // 故障标志，本件结构性不置位 / fault flag, never raised by this component
    bValid      : BOOL;     // 结果可用标志 / result usable flag
END_VAR
VAR CONSTANT
    DL_TEN      : UDINT := 10;              // 十进制基数 [无量纲] / decimal radix, dimensionless
    DL_ONE      : UDINT := 1;               // 整数一，零值也占一位 [位] / integer one, zero still occupies one digit [digit]
    DL_LOOP_MAX : UDINT := 10;              // 循环上界，等于最大位数 [位] / loop cap equal to the largest width [digit]
END_VAR
VAR
    nRest       : UDINT;    // 降位过程中的剩余值 / remaining value while descending
    nDigits     : UDINT;    // 已计位数 / digits counted so far
    nGuard      : UDINT;    // 循环守卫计数 / loop guard counter
END_VAR

// 段 1｜出口预置：零值占一位，故计数从 1 起 / segment 1, preset with one digit because zero occupies one position
FC_DL_IntDigitCountUdint := 0;  // 缺省 0 / default zero
eErr    := 0;                   // 零码位范式 / zero-code rule
bError  := FALSE;               // 本件不产生故障级 / this component raises no fault
bValid  := TRUE;                // 全定义域恒可完成 / always completes over the whole domain
nRest   := nVal;                // 从输入起步 / start from the input
nDigits := DL_ONE;              // 零值即一位 / zero already occupies one digit
nGuard  := 0;                   // 守卫清零 / clear the guard

// 段 2｜降位：剩余值 ≥ 10 才进一位 / segment 2, divide down while the remainder is ten or more
WHILE (nRest >= DL_TEN) AND (nGuard < DL_LOOP_MAX) DO
    nGuard  := nGuard + DL_ONE;         // 守卫自增 / advance the guard
    nRest   := nRest / DL_TEN;          // 降一位 / shift one digit down
    nDigits := nDigits + DL_ONE;        // 位数加一 / one more digit
END_WHILE

// 段 3｜出口 / segment 3, exit
FC_DL_IntDigitCountUdint := nDigits;    // 1~10 / one to ten
END_FUNCTION

(* ---- FC_DL_IntDigitSumUdint.st ---- *)
(*==============================================================================
 * 组件名称 : FC_DL_IntDigitSumUdint ｜ 子库 : DL_MathData ｜ v1.0.0 ｜ 2026-11-24
 * 平台     : CODESYS 3.5 / TwinCAT 3 / InoProShop / Machine Expert（纯 IEC，无厂商库）
 * 功能简介 : 无符号整数的十进制各位数字之和（数字根母函数）。逐次取余取位再整除降位，
 *            纯整数实现，禁字符串转换（字符串转换在多平台补零/符号口径不一致）。
 * 契约     : 返回各位数字之和（最大 10 位 × 9 = 90）；nVal = 0 返回 0。
 *            循环次数以 nVal 位数为上界，结构性有限。
 * 依赖     : 无 DL_ 内部依赖（R16 自足实现），无标准库函数调用
 * 错误码   : R297 零码位范式：eErr 恒 0，仅以 bError / bValid 表达（本件结构性不置 bError）
 * 红线自检 : R1 零全局 R2 零%I/%Q R3 纯IEC R4 除数为常量 10、循环上界固定
 *            R5 双语注释 R6 N/A（无状态机）R7 N/A（无定时器/沿实例）
 *            R10 无类型转换 R11 全声明行分号 R15 标识符零保留字冲突 R18 N/A（无 bReset）
 * 修订历史 : 2026-11-24 R79-A 首版（整数数论族 3/8）
 *============================================================================*)
FUNCTION FC_DL_IntDigitSumUdint : UDINT
VAR_INPUT
    nVal        : UDINT;    // 被分解整数，全域 0~16#FFFF_FFFF [无量纲] / value to decompose over the whole unsigned range
END_VAR
VAR_OUTPUT
    eErr        : UDINT;    // 错误码，零码位范式恒 0 / error id, always zero under the zero-code rule
    bError      : BOOL;     // 故障标志，本件结构性不置位 / fault flag, never raised by this component
    bValid      : BOOL;     // 结果可用标志 / result usable flag
END_VAR
VAR CONSTANT
    DL_TEN      : UDINT := 10;              // 十进制基数 [无量纲] / decimal radix, dimensionless
    DL_ZERO     : UDINT := 0;               // 整数零哨兵 [无量纲] / integer zero sentinel, dimensionless
    DL_LOOP_MAX : UDINT := 10;              // UDINT 十进制最大位数，循环上界 [位] / largest decimal width of an unsigned value [digit]
END_VAR
VAR
    nRest       : UDINT;    // 降位过程中的剩余值 / remaining value while descending
    nSum        : UDINT;    // 各位数字累计和 / accumulated digit sum
    nGuard      : UDINT;    // 循环守卫计数，防遍历失控 / loop guard counter
END_VAR

// 段 1｜出口预置 / segment 1, preset the exit
FC_DL_IntDigitSumUdint := 0;    // 缺省 0 / default zero
eErr   := 0;                    // 零码位范式 / zero-code rule
bError := FALSE;                // 本件不产生故障级 / this component raises no fault
bValid := TRUE;                 // 分解对全定义域恒可完成 / the decomposition always completes over the whole domain
nRest  := nVal;                 // 从输入起步 / start from the input
nSum   := DL_ZERO;              // 累计清零 / clear the accumulator
nGuard := DL_ZERO;              // 守卫清零 / clear the guard

// 段 2｜逐位取余累加，整除降位；剩余为 0 即停 / segment 2, take the remainder, add it, divide down
WHILE (nRest <> DL_ZERO) AND (nGuard < DL_LOOP_MAX) DO
    nGuard := nGuard + 1;                       // 守卫自增 / advance the guard
    nSum   := nSum + (nRest MOD DL_TEN);        // 取个位并累加 / take the units digit and accumulate
    nRest  := nRest / DL_TEN;                   // 降一位 / shift one digit down
END_WHILE

// 段 3｜出口 / segment 3, exit
FC_DL_IntDigitSumUdint := nSum;                 // 各位数字之和 / the digit sum
END_FUNCTION

(* ---- FC_DL_InterpolateTable2D.st ---- *)
(*
    FC_DL_InterpolateTable2D —— 二维标定表双线性插值
    ------------------------------------------------------------------
    分类      : DL_MathData / Interpolate
    前缀      : FC_DL_
    版本      : 1.0.0
    溯源      : T2-1 LGF · Math（只借「标度 / 插值属 Math 组」的分类事实与参数域组织
                方式；双线性公式为公开数学，实现、码位、行主序约定 100% 自有）；
                clean-room 重写，未复制任何闭源厂商源码，参考实现仅限 MIT/Apache 许可
    平台      : 纯 IEC 61131-3，CODESYS V3.5+ / TwinCAT 3 / InoProShop 通用
    作者      : 道莅代码库 · PLC编程专家（R18）
    ------------------------------------------------------------------
    功能说明  : 8x8 标定网格上做双线性插值，典型场景：温度—压力二维补偿表、
                阀门流量特性双参数表、视觉标定畸变修正；库内 MultiPointLinear 只做
                一维，二维场景现场长期靠梯形图硬编码，本件即补此缺口；
                防御链：点数闸 → 网格严格递增校验 → 坐标非有限闸 → 退化格防除零闸
                → 索引上界闸 → 结果非有限复检，每一闸都在索引或除法之前；
                定位用线性扫描（点数不超过 8，避免二分的边界 off-by-one），
                值表按行主序一维存放，不用多维数组规避平台差异。
    错误码    : 16#0001_023F 输入落网格外已钳位，或遇退化格（跨度约等于 0）按该角值直取——信息级，正常防御
                16#0001_0240 预留禁用（信息级，不得挪用）
                16#0001_0315 点数或网格非法（越界、非严格递增）——故障级，返回首值
                16#0001_0316 插值坐标或结果非有限（NaN / 正负 INF）——故障级，返回首值
                16#0001_0317 预留禁用（故障级，不得挪用）
    码位总账  : 16#0001_023F 用 / 16#0001_0240 预留 ｜ 16#0001_0315 用 / 16#0001_0316 用 / 16#0001_0317 预留
    状态机    : N/A —— 纯函数无顺序状态机，无 CASE 可写，非法状态不可能出现
    采样约定  : 纯组合函数，无定时器、无内部驻留状态；网格与值表由调用方保证
                在调用拍内不被并发改写（本库统一约定：标定表只在停机态下发）。
    修订记录  : 2026-11-16 v1.0.0 首次入库（R18）
*)
FUNCTION FC_DL_InterpolateTable2D : REAL
VAR_INPUT
    afGridX      : ARRAY[0..7] OF REAL;        // X 轴网格，必须严格递增，有效项 0~uCountX-1 [用户单位] / X grid, strictly increasing, valid items 0~uCountX-1 [user unit]
    afGridY      : ARRAY[0..7] OF REAL;        // Y 轴网格，必须严格递增，有效项 0~uCountY-1 [用户单位] / Y grid, strictly increasing, valid items 0~uCountY-1 [user unit]
    afValue      : ARRAY[0..63] OF REAL;       // 值表，行主序：索引 = nIy * uCountX + nIx [用户单位] / value table, row major, index = nIy * uCountX + nIx [user unit]
    uCountX      : UINT := 2;                  // X 有效点数 [点]，范围 2~8 / valid X point count [pt], range 2~8
    uCountY      : UINT := 2;                  // Y 有效点数 [点]，范围 2~8 / valid Y point count [pt], range 2~8
    fX           : REAL := 0.0;                // 待插值 X [用户单位] / X to interpolate [user unit]
    fY           : REAL := 0.0;                // 待插值 Y [用户单位] / Y to interpolate [user unit]
    bExtrapolate : BOOL := FALSE;              // FALSE 边界钳位（推荐）/ TRUE 单格外延 / FALSE clamps at the border, TRUE extrapolates one cell
END_VAR
VAR_OUTPUT
    eErr       : UDINT;                        // 错误码，0=正常 / error id, 0=ok
    bError     : BOOL;                         // 故障标志，eErr 为故障级时 TRUE / error flag, TRUE on fault-level eErr
    bValid     : BOOL;                         // 结果是否可用 / result usable flag
    bOutOfGrid : BOOL;                         // 输入落在网格外（钳位或外延生效）/ input falls outside the grid (clamp or extrapolation applied)
END_VAR
VAR
    uIx      : UINT;                           // X 网格遍历游标 [点] / X grid traversal cursor [pt]
    uIy      : UINT;                           // Y 网格遍历游标 [点] / Y grid traversal cursor [pt]
    uIxSel   : UINT;                           // 命中的 X 单元下界序号 [点] / selected lower X cell index [pt]
    uIySel   : UINT;                           // 命中的 Y 单元下界序号 [点] / selected lower Y cell index [pt]
    uBase    : UINT;                           // 四角首索引（行主序）[无量纲] / first corner index in row major order [dimensionless]
    uIdx11   : UINT;                           // 对角索引 uIdx11，用于上界闸 [无量纲] / diagonal index used by the upper bound gate [dimensionless]
    fTx      : REAL;                           // X 方向归一化插值系数 0~1 / normalised interpolation factor along X, 0~1
    fTy      : REAL;                           // Y 方向归一化插值系数 0~1 / normalised interpolation factor along Y, 0~1
    fV00     : REAL;                           // 左下角值 [用户单位] / lower left corner value [user unit]
    fV10     : REAL;                           // 右下角值 [用户单位] / lower right corner value [user unit]
    fV01     : REAL;                           // 左上角值 [用户单位] / upper left corner value [user unit]
    fV11     : REAL;                           // 右上角值 [用户单位] / upper right corner value [user unit]
    fSpanX   : REAL;                           // X 单元跨度 [用户单位] / X cell span [user unit]
    fSpanY   : REAL;                           // Y 单元跨度 [用户单位] / Y cell span [user unit]
    fRes     : REAL;                           // 插值结果中间量 [用户单位] / interpolation result intermediate [user unit]
    bFoundX  : BOOL;                           // X 定位命中标志 / X location found flag
    bFoundY  : BOOL;                           // Y 定位命中标志 / Y location found flag
    bNonFin  : BOOL;                           // 非有限判定中间标志 / non-finite detection intermediate flag
END_VAR
VAR CONSTANT
    DL_2D_MAX        : UINT := 8;              // 单轴点数上限 [点] / per axis point upper bound [pt]
    DL_2D_CELLS      : UINT := 64;             // 值表容量 [个] / value table capacity [item]
    DL_2D_LAST_CELL  : UINT := 63;             // 值表末索引 [个] / last value table index [item]
    DL_FLOAT_EPS     : REAL := 1.0E-6;         // 浮点判等容差 [无量纲] / float equality tolerance [dimensionless]
    DL_2D_INF_GUARD  : REAL := 4.0E38;         // 非有限幅值判定阈值，高于 REAL 最大有限值 [用户单位] / non-finite magnitude guard above the largest finite REAL [user unit]
    DL_2D_ONE        : REAL := 1.0;            // 归一化上界与补数基数 [无量纲] / normalisation upper bound and complement base [dimensionless]
    DL_2D_ZERO       : REAL := 0.0;            // 零值常量，避免裸字面量 [无量纲] / zero constant, avoids a bare literal [dimensionless]
END_VAR

// 段 1｜返回值与错误状态预置 / segment 1, preset return value and error status
FC_DL_InterpolateTable2D := DL_2D_ZERO;        // 故障缺省返回 0 / fault default returns zero
eErr := 0;                                     // 预置无错误 / preset no error
bError := FALSE;                               // 预置无故障 / preset no fault
bValid := FALSE;                               // 预置结果不可用 / preset unusable
bOutOfGrid := FALSE;                           // 预置落在网格内 / preset inside the grid

// 段 2｜点数闸：先判界再索引，绝不越界读数组 / segment 2, point count gate before any indexing
IF (uCountX < 2) OR (uCountX > DL_2D_MAX) OR (uCountY < 2) OR (uCountY > DL_2D_MAX) THEN
    eErr := 16#0001_0315;                      // 点数非法故障码 / illegal point count fault id
    bError := TRUE;                            // 置故障标志 / raise the error flag
    FC_DL_InterpolateTable2D := afValue[0];    // 返回首值，索引 0 恒存在 / return the first value, index zero always exists
    RETURN;                                    // 故障级提前返回 / early return on fault
END_IF

// 段 3｜坐标非有限闸（NaN 自不等 + 幅值判正负 INF）/ segment 3, non-finite coordinate gate
bNonFin := (fX <> fX) OR (fX > DL_2D_INF_GUARD) OR (fX < -DL_2D_INF_GUARD)
        OR (fY <> fY) OR (fY > DL_2D_INF_GUARD) OR (fY < -DL_2D_INF_GUARD); // 非有限综合判定 / combined non-finite check
IF bNonFin THEN
    eErr := 16#0001_0316;                      // 坐标非有限故障码 / non-finite coordinate fault id
    bError := TRUE;                            // 置故障标志 / raise the error flag
    FC_DL_InterpolateTable2D := afValue[0];    // 返回首值 / return the first value
    RETURN;                                    // 故障级提前返回 / early return on fault
END_IF

// 段 4｜网格严格递增校验（用大于号逐点比较，禁用浮点判等）/ segment 4, strict monotonic grid check
FOR uIx := 1 TO uCountX - 1 DO
    IF NOT (afGridX[uIx] > afGridX[uIx - 1]) THEN
        eErr := 16#0001_0315;                  // 网格非严格递增故障码 / non monotonic grid fault id
        bError := TRUE;                        // 置故障标志 / raise the error flag
        FC_DL_InterpolateTable2D := afValue[0];// 返回首值 / return the first value
        RETURN;                                // 故障级提前返回 / early return on fault
    END_IF
END_FOR
FOR uIy := 1 TO uCountY - 1 DO
    IF NOT (afGridY[uIy] > afGridY[uIy - 1]) THEN
        eErr := 16#0001_0315;                  // Y 网格非严格递增故障码 / non monotonic Y grid fault id
        bError := TRUE;                        // 置故障标志 / raise the error flag
        FC_DL_InterpolateTable2D := afValue[0];// 返回首值 / return the first value
        RETURN;                                // 故障级提前返回 / early return on fault
    END_IF
END_FOR

// 段 5｜线性扫描定位单元（上界 uCountX-2，避免 off-by-one）/ segment 5, linear cell location
uIxSel := 0;                                   // 默认落最低单元 / default to the lowest cell
bFoundX := FALSE;                              // 命中标志先清 / clear the found flag
FOR uIx := 0 TO uCountX - 2 DO
    IF (NOT bFoundX) AND (fX <= afGridX[uIx + 1]) THEN
        uIxSel := uIx;                         // 命中第一个上界不小于输入的单元 / the first cell whose upper bound is not below the input
        bFoundX := TRUE;                       // 命中即锁定，后续不再覆盖 / lock the hit, later cells never overwrite it
    END_IF
END_FOR
IF NOT bFoundX THEN
    uIxSel := uCountX - 2;                     // 高于网格顶，取最高单元 / above the top, take the highest cell
    bOutOfGrid := TRUE;                        // 标记落在网格外 / flag the out-of-grid input
END_IF
IF fX < afGridX[0] THEN
    uIxSel := 0;                               // 低于网格底，取最低单元 / below the bottom, take the lowest cell
    bOutOfGrid := TRUE;                        // 标记落在网格外 / flag the out-of-grid input
END_IF
uIySel := 0;                                   // 默认落最低单元 / default to the lowest cell
bFoundY := FALSE;                              // 命中标志先清 / clear the found flag
FOR uIy := 0 TO uCountY - 2 DO
    IF (NOT bFoundY) AND (fY <= afGridY[uIy + 1]) THEN
        uIySel := uIy;                         // 命中第一个上界不小于输入的单元 / the first cell whose upper bound is not below the input
        bFoundY := TRUE;                       // 命中即锁定 / lock the hit
    END_IF
END_FOR
IF NOT bFoundY THEN
    uIySel := uCountY - 2;                     // 高于网格顶，取最高单元 / above the top, take the highest cell
    bOutOfGrid := TRUE;                        // 标记落在网格外 / flag the out-of-grid input
END_IF
IF fY < afGridY[0] THEN
    uIySel := 0;                               // 低于网格底，取最低单元 / below the bottom, take the lowest cell
    bOutOfGrid := TRUE;                        // 标记落在网格外 / flag the out-of-grid input
END_IF

// 段 6｜退化格防除零：跨度绝对值不大于容差时不除，系数取 0 按该角值直取 / segment 6, degenerate cell division guard
fSpanX := afGridX[uIxSel + 1] - afGridX[uIxSel]; // X 单元跨度 / X cell span
IF ABS(fSpanX) <= DL_FLOAT_EPS THEN
    fTx := DL_2D_ZERO;                         // 跨度近零，系数取 0，绝不除 / span near zero, factor zero, no division
    eErr := 16#0001_023F;                      // 退化格提示（信息级不置故障）/ degenerate cell hint, info level never raises a fault
ELSE
    fTx := (fX - afGridX[uIxSel]) / fSpanX;    // 除号在防零闸之后 / the division happens after the guard
END_IF
fSpanY := afGridY[uIySel + 1] - afGridY[uIySel]; // Y 单元跨度 / Y cell span
IF ABS(fSpanY) <= DL_FLOAT_EPS THEN
    fTy := DL_2D_ZERO;                         // 跨度近零，系数取 0 / span near zero, factor zero
    eErr := 16#0001_023F;                      // 退化格提示（信息级不置故障）/ degenerate cell hint, info level never raises a fault
ELSE
    fTy := (fY - afGridY[uIySel]) / fSpanY;    // 除号在防零闸之后 / the division happens after the guard
END_IF

// 段 7｜边界策略：钳位（推荐）或单格外延 / segment 7, border policy, clamp or single cell extrapolation
IF bExtrapolate THEN
    IF bOutOfGrid THEN
        eErr := 16#0001_023F;                  // 外延生效提示（信息级不置故障）/ extrapolation hint, info level never raises a fault
    END_IF
ELSE
    IF fTx < DL_2D_ZERO THEN
        fTx := DL_2D_ZERO;                     // 下侧钳位 / clamp on the low side
        bOutOfGrid := TRUE;                    // 标记落网格外 / flag the out-of-grid input
    END_IF
    IF fTx > DL_2D_ONE THEN
        fTx := DL_2D_ONE;                      // 上侧钳位 / clamp on the high side
        bOutOfGrid := TRUE;                    // 标记落网格外 / flag the out-of-grid input
    END_IF
    IF fTy < DL_2D_ZERO THEN
        fTy := DL_2D_ZERO;                     // 下侧钳位 / clamp on the low side
        bOutOfGrid := TRUE;                    // 标记落网格外 / flag the out-of-grid input
    END_IF
    IF fTy > DL_2D_ONE THEN
        fTy := DL_2D_ONE;                      // 上侧钳位 / clamp on the high side
        bOutOfGrid := TRUE;                    // 标记落网格外 / flag the out-of-grid input
    END_IF
    IF bOutOfGrid THEN
        eErr := 16#0001_023F;                  // 钳位生效提示（信息级不置故障）/ clamp hint, info level never raises a fault
    END_IF
END_IF

// 段 8｜四角索引上界闸：一切索引在取用前判界 / segment 8, corner index upper bound gate
uBase := uIySel * uCountX + uIxSel;            // 行主序首索引 / first corner index in row major order
uIdx11 := uBase + uCountX + 1;                 // 对角索引 / diagonal index
IF uIdx11 > DL_2D_LAST_CELL THEN
    eErr := 16#0001_0315;                      // 索引越界故障码 / index out of range fault id
    bError := TRUE;                            // 置故障标志 / raise the error flag
    FC_DL_InterpolateTable2D := afValue[0];    // 返回首值 / return the first value
    RETURN;                                    // 故障级提前返回 / early return on fault
END_IF
fV00 := afValue[uBase];                        // 左下角值 / lower left value
fV10 := afValue[uBase + 1];                    // 右下角值 / lower right value
fV01 := afValue[uBase + uCountX];              // 左上角值 / upper left value
fV11 := afValue[uIdx11];                       // 右上角值 / upper right value

// 段 9｜双线性合成 / segment 9, bilinear composition
fRes := fV00 * (DL_2D_ONE - fTx) * (DL_2D_ONE - fTy)
      + fV10 * fTx * (DL_2D_ONE - fTy)
      + fV01 * (DL_2D_ONE - fTx) * fTy
      + fV11 * fTx * fTy;                      // 四角加权求和 / weighted sum of the four corners
bNonFin := (fRes <> fRes) OR (fRes > DL_2D_INF_GUARD) OR (fRes < -DL_2D_INF_GUARD); // 结果非有限复检 / result non-finite recheck
IF bNonFin THEN
    eErr := 16#0001_0316;                      // 结果非有限故障码 / non-finite result fault id
    bError := TRUE;                            // 置故障标志 / raise the error flag
    FC_DL_InterpolateTable2D := afValue[0];    // 返回首值 / return the first value
    RETURN;                                    // 故障级提前返回 / early return on fault
END_IF

// 段 10｜出口 / segment 10, exit
FC_DL_InterpolateTable2D := fRes;              // 输出插值结果 / publish the interpolated result
bValid := TRUE;                                // 结果可用 / the result is usable
END_FUNCTION

(* ---- FC_DL_InterpolateTable3D.st ---- *)
(*
  ==================================================================
  组件名 Component  : FC_DL_InterpolateTable3D
  分类   Category   : DL_MathData
  复杂度 Complexity  : 高
  版本   Version    : 1.0.1
  功能   Purpose    : 三维表三线性插值。三条轴向量（升序）定位所在单元，索引钳位到
                      [0, n-2]，单元内按 X→Y→Z 三次线性插值出结果；轴乱序、
                      输入非有限、表值非有限三类异常各自置码并拒绝出值。
  来源   Source     : t2-1-lgf-math（LGF Math 插值族三维变体）
  溯源   Origin     : 三线性插值属公开数值语义，clean-room 自研实现，未复制 LGF
                      或任何厂商私有库源码。
  平台   Platform   : 纯 IEC 61131-3（FOR / 四则运算 / ABS），三平台通用
  分工声明 Split     : 与 FC_DL_InterpolateTable2D（2D 属主）与 FB_DL_LineInterp2Axis
                      （轴对直线插值）分工——本件为三维表族谱最高维成员，只做
                      三线性单元插值，不做二维降维代理、不做外插。
  作者   Author     : 道莅代码库 · PLC 编程专家（R60）
  ------------------------------------------------------------------
  边界 Boundary     :
                      一 轴向量必须严格升序（aX[i] < aX[i+1]）：非升序判故障级码并
                         拒绝插值，不做排序修正（改调用方数据属越界，边界五）；
                      二 单元索引钳位到 [0, n-2]：输入低于首节点落单元 0、高于末节点
                         落单元 n-2（外插不外推，等价于边界保持）；
                      三 有限性闸覆盖参与换算的每个浮点引脚（R272 自证）：标量
                         fX / fY / fZ 逐个点名，轴向量与表值按参与元素逐个判；
                      四 结果非有限兜底同拍置 eErr + bError + bValid 三件套（R258）；
                      五 只读轴向量与表数组，不改调用方数据（PercentileLReal 纪律）。
  错误码   Codes    :
    16#0001_0626【信息级】轴元素数越域已钳位（<2 或 >16）
    16#0001_0627【故障级】轴向量非严格升序，拒绝插值
    16#0001_0628【故障级】输入坐标含非有限值，拒绝插值
    16#0001_0629【故障级】轴或表值含非有限值，拒绝插值
    16#0001_0630【故障级】插值结果非有限（复检兜底，R190 独立码）
  验收   Acceptance :
    算法已证（脚本）：未跑 ｜ 编译器已证（三平台）：未跑
    V1 轴 0/10、表值仅随 X 线性（f=2X）→ 输入 (5,0,0) 得 10.0
    V2 输入 (20,0,0) 高于末节点 → 落末单元，得末节点值（不外推）
    V3 aX = 0/10/5（乱序）→ 码 0627、bValid = FALSE
    V4 fX = NaN → 码 0628、bValid = FALSE、fOut = 0
  修订记录 Revision  :
    2026-11-21  v1.0.0  R60 首版（批 3 · 序号 9）
    2026-11-21  v1.0.1  R61 返修：D3 三轴向量逐元素非有限点名（R272 全量）；
                        D4 信息级 0626 两处不再置 bError（R285 口径统一）；
                        D8 段 6 八角点判缩进对齐；D9 新增 0630 结果非有限码
  ==================================================================
*)
FUNCTION FC_DL_InterpolateTable3D : LREAL
VAR_IN_OUT
    afX     : ARRAY[0..15] OF LREAL;             // X 轴向量（严格升序）[用户单位] / the X axis vector, strictly ascending
    afY     : ARRAY[0..15] OF LREAL;             // Y 轴向量（严格升序）[用户单位] / the Y axis vector, strictly ascending
    afZ     : ARRAY[0..15] OF LREAL;             // Z 轴向量（严格升序）[用户单位] / the Z axis vector, strictly ascending
    afTable : ARRAY[0..15, 0..15, 0..15] OF LREAL; // 表值 [工程单位]，维序 X,Y,Z / the table values with the dimension order X, Y, Z
END_VAR
VAR_INPUT
    nX : DINT;   // X 轴元素数 [个]，合法域 2..16 / the X element count, legal from two to sixteen
    nY : DINT;   // Y 轴元素数 [个]，合法域 2..16 / the Y element count, legal from two to sixteen
    nZ : DINT;   // Z 轴元素数 [个]，合法域 2..16 / the Z element count, legal from two to sixteen
    fX : LREAL;  // X 输入坐标 [用户单位] / the X input coordinate
    fY : LREAL;  // Y 输入坐标 [用户单位] / the Y input coordinate
    fZ : LREAL;  // Z 输入坐标 [用户单位] / the Z input coordinate
END_VAR
VAR_OUTPUT
    bValid : BOOL;  // 结果可用标志 [-] / the result usable flag
    eErr   : UDINT; // 错误码，0 = 正常 / the error code, zero is ok
    bError : BOOL;  // 错误标志，eErr 非 0 时为真 / the error flag, true when eErr is nonzero
END_VAR
VAR
    nIx     : DINT;  // X 单元索引 [下标] / the X cell index
    nIy     : DINT;  // Y 单元索引 [下标] / the Y cell index
    nIz     : DINT;  // Z 单元索引 [下标] / the Z cell index
    k       : DINT;  // 轴遍历索引 [下标] / the axis loop index
    nUseX   : DINT;  // 钳位后 X 元素数 [个] / the clamped X count
    nUseY   : DINT;  // 钳位后 Y 元素数 [个] / the clamped Y count
    nUseZ   : DINT;  // 钳位后 Z 元素数 [个] / the clamped Z count
    fTx     : LREAL; // X 单元内归一化位置 [-] / the normalised X position inside the cell
    fTy     : LREAL; // Y 单元内归一化位置 [-] / the normalised Y position inside the cell
    fTz     : LREAL; // Z 单元内归一化位置 [-] / the normalised Z position inside the cell
    fSpan   : LREAL; // 单元宽度工作副本 [用户单位] / the cell span copy
    fC000   : LREAL; // 角点 (i,j,k) 表值 [工程单位] / the corner value at i, j, k
    fC100   : LREAL; // 角点 (i+1,j,k) 表值 [工程单位] / the corner value at i plus one, j, k
    fC010   : LREAL; // 角点 (i,j+1,k) 表值 [工程单位] / the corner value at i, j plus one, k
    fC110   : LREAL; // 角点 (i+1,j+1,k) 表值 [工程单位] / the corner value at i plus one, j plus one, k
    fC001   : LREAL; // 角点 (i,j,k+1) 表值 [工程单位] / the corner value at i, j, k plus one
    fC101   : LREAL; // 角点 (i+1,j,k+1) 表值 [工程单位] / the corner value at i plus one, j, k plus one
    fC011   : LREAL; // 角点 (i,j+1,k+1) 表值 [工程单位] / the corner value at i, j plus one, k plus one
    fC111   : LREAL; // 角点 (i+1,j+1,k+1) 表值 [工程单位] / the corner value at i plus one, j plus one, k plus one
    fX0     : LREAL; // 单元 X 下节点坐标 [用户单位] / the cell lower X node
    fY0     : LREAL; // 单元 Y 下节点坐标 [用户单位] / the cell lower Y node
    fZ0     : LREAL; // 单元 Z 下节点坐标 [用户单位] / the cell lower Z node
    fA0     : LREAL; // X 向插值低端结果（k 层）[工程单位] / the X interpolation at the lower Z layer
    fA1     : LREAL; // X 向插值低端结果（k+1 层）[工程单位] / the X interpolation at the upper Z layer
    fB0     : LREAL; // Y 向插值结果（k 层）[工程单位] / the Y interpolation at the lower Z layer
    fB1     : LREAL; // Y 向插值结果（k+1 层）[工程单位] / the Y interpolation at the upper Z layer
    bClamp  : BOOL;  // 元素数钳位标记 [-] / the element count clamp flag
    bOrder  : BOOL;  // 轴乱序标记 [-] / the axis order fault flag
    bNonFin : BOOL;  // 非有限标记 [-] / the non finite flag
END_VAR
VAR CONSTANT
    DL_I3D_NMAX : DINT := 16; // 轴元素容量上界 [个]，与数组第一维一致 / the axis capacity aligned with the first dimension
    DL_I3D_TOL  : LREAL := 1.0E-12; // 差值比较容差 [用户单位] / the difference comparison tolerance
END_VAR

// 段 1｜返回值与错误状态预置安全值（四段式第一段，R45）+ 局部量显式预置（R254）/ segment 1, the preset of the return, the codes and the local guards
FC_DL_InterpolateTable3D := 0.0; // 返回值预置安全值零 / preset the return to zero
bValid := FALSE; // 有效标志预置假 / preset the validity false
eErr := 16#0000_0000; // 错误码预置正常 / preset the code to ok
bError := FALSE; // 错误标志预置假 / preset the error flag false
bClamp := FALSE; // 钳位标记预置假 / preset the clamp flag false
bOrder := FALSE; // 乱序标记预置假 / preset the order fault flag false
bNonFin := FALSE; // 非有限标记预置假 / preset the non finite flag false
nIx := 0; // X 单元索引预置零 / preset the X cell index zero
nIy := 0; // Y 单元索引预置零 / preset the Y cell index zero
nIz := 0; // Z 单元索引预置零 / preset the Z cell index zero
fTx := 0.0; // X 归一化位置预置零 / preset the X position zero
fTy := 0.0; // Y 归一化位置预置零 / preset the Y position zero
fTz := 0.0; // Z 归一化位置预置零 / preset the Z position zero
fSpan := 0.0; // 单元宽度预置零 / preset the cell span zero
fX0 := 0.0; // X 下节点预置零 / preset the X lower node zero
fY0 := 0.0; // Y 下节点预置零 / preset the Y lower node zero
fZ0 := 0.0; // Z 下节点预置零 / preset the Z lower node zero

// 段 2｜元素数域闸（<2 早退，>16 钳位，边界二）/ segment 2, the element count gate
IF (nX < 2) OR (nY < 2) OR (nZ < 2) THEN // 任轴少于两个节点，无单元可插值 / fewer than two nodes leave no cell
    eErr := 16#0001_0626; // 信息级：轴元素数越域已钳位（信息级不置 bError，R285 口径统一）/ informational, the element count clamped, no fault bit by the unified grade rule
    RETURN; // 早退 / early return
END_IF
nUseX := nX; // X 元素数域内接管 / take the X count
nUseY := nY; // Y 元素数域内接管 / take the Y count
nUseZ := nZ; // Z 元素数域内接管 / take the Z count
IF nUseX > DL_I3D_NMAX THEN // 超容量 / above the capacity
    nUseX := DL_I3D_NMAX; // 钳到容量 / clamp to the capacity
    bClamp := TRUE; // 置钳位标记 / raise the clamp flag
END_IF
IF nUseY > DL_I3D_NMAX THEN // 超容量 / above the capacity
    nUseY := DL_I3D_NMAX; // 钳到容量 / clamp to the capacity
    bClamp := TRUE; // 置钳位标记 / raise the clamp flag
END_IF
IF nUseZ > DL_I3D_NMAX THEN // 超容量 / above the capacity
    nUseZ := DL_I3D_NMAX; // 钳到容量 / clamp to the capacity
    bClamp := TRUE; // 置钳位标记 / raise the clamp flag
END_IF
IF bClamp THEN // 钳位置信息级 / raise the informational code on a clamp
    eErr := 16#0001_0626; // 信息级：轴元素数越域已钳位 / informational, the element count clamped
    bError := TRUE; // 置错误标志 / raise the error flag
END_IF

// 段 3｜轴严格升序与有限性闸（轴与输入坐标，边界一三）/ segment 3, the axis order and the finiteness gate
FOR k := 0 TO nUseX - 2 DO // X 轴相邻比较 / the X neighbour comparison
    IF (afX[k] <> afX[k]) OR ((afX[k] - afX[k]) <> (afX[k] - afX[k]))
    OR (afX[k + 1] <> afX[k + 1]) OR ((afX[k + 1] - afX[k + 1]) <> (afX[k + 1] - afX[k + 1])) THEN // X 轴相邻元素逐个非有限判（D3 返修，R272 点名）/ the adjacent X elements tested for finiteness one by one
        bNonFin := TRUE; // 置非有限标记 / raise the non finite flag
    END_IF
    IF afX[k] >= afX[k + 1] THEN // 非严格升序 / not strictly ascending
        bOrder := TRUE; // 置乱序标记 / raise the order flag
    END_IF
END_FOR
FOR k := 0 TO nUseY - 2 DO // Y 轴相邻比较 / the Y neighbour comparison
    IF (afY[k] <> afY[k]) OR ((afY[k] - afY[k]) <> (afY[k] - afY[k]))
    OR (afY[k + 1] <> afY[k + 1]) OR ((afY[k + 1] - afY[k + 1]) <> (afY[k + 1] - afY[k + 1])) THEN // Y 轴相邻元素逐个非有限判（D3 返修）/ the adjacent Y elements tested for finiteness
        bNonFin := TRUE; // 置非有限标记 / raise the non finite flag
    END_IF
    IF afY[k] >= afY[k + 1] THEN // 非严格升序 / not strictly ascending
        bOrder := TRUE; // 置乱序标记 / raise the order flag
    END_IF
END_FOR
FOR k := 0 TO nUseZ - 2 DO // Z 轴相邻比较 / the Z neighbour comparison
    IF (afZ[k] <> afZ[k]) OR ((afZ[k] - afZ[k]) <> (afZ[k] - afZ[k]))
    OR (afZ[k + 1] <> afZ[k + 1]) OR ((afZ[k + 1] - afZ[k + 1]) <> (afZ[k + 1] - afZ[k + 1])) THEN // Z 轴相邻元素逐个非有限判（D3 返修）/ the adjacent Z elements tested for finiteness
        bNonFin := TRUE; // 置非有限标记 / raise the non finite flag
    END_IF
    IF afZ[k] >= afZ[k + 1] THEN // 非严格升序 / not strictly ascending
        bOrder := TRUE; // 置乱序标记 / raise the order flag
    END_IF
END_FOR
IF bNonFin THEN // 轴向量含非有限（NaN 使序闸恒假，须先于乱序判拒算，D3）/ a non finite axis element, gated ahead of the order test
    eErr := 16#0001_0629; // 故障级：轴或表值含非有限值 / fault grade, a non finite axis or table value
    bError := TRUE; // 置错误标志（R45 配对）/ raise the error flag, paired with the fault code
    bValid := FALSE; // 结果不可用 / the result void
    RETURN; // 早退 / early return
END_IF
IF bOrder THEN // 轴乱序即拒算（不排序修正，边界一）/ refuse on a disorder, no sorting
    eErr := 16#0001_0627; // 故障级：轴向量非严格升序 / fault grade, the axis is not strictly ascending
    bError := TRUE; // 置错误标志（R45 配对）/ raise the error flag, paired with the fault code
    bValid := FALSE; // 结果不可用 / the result void
    RETURN; // 早退 / early return
END_IF
IF (fX <> fX) OR ((fX - fX) <> (fX - fX)) OR (fY <> fY) OR ((fY - fY) <> (fY - fY))
OR (fZ <> fZ) OR ((fZ - fZ) <> (fZ - fZ)) THEN // 三个输入坐标逐个非有限判（R272 点名）/ the three input coordinates tested one by one
    eErr := 16#0001_0628; // 故障级：输入坐标含非有限值 / fault grade, a non finite input coordinate
    bError := TRUE; // 置错误标志（R45 配对）/ raise the error flag, paired with the fault code
    bValid := FALSE; // 结果不可用 / the result void
    RETURN; // 早退 / early return
END_IF

// 段 4｜三轴单元定位（线性查找 + 钳位到 [0, n-2]，输入不外推）/ segment 4, the cell location clamped to the legal index band
nIx := 0; // X 单元索引从零起 / the X index starts at zero
FOR k := 0 TO nUseX - 2 DO // 升序轴线性定位 / the linear location on an ascending axis
    IF fX >= afX[k] THEN // 已过该下节点 / the input is past this lower node
        nIx := k; // 记录候选单元 / register the candidate cell
    END_IF
END_FOR
nIy := 0; // Y 单元索引从零起 / the Y index starts at zero
FOR k := 0 TO nUseY - 2 DO // 升序轴线性定位 / the linear location on an ascending axis
    IF fY >= afY[k] THEN // 已过该下节点 / the input is past this lower node
        nIy := k; // 记录候选单元 / register the candidate cell
    END_IF
END_FOR
nIz := 0; // Z 单元索引从零起 / the Z index starts at zero
FOR k := 0 TO nUseZ - 2 DO // 升序轴线性定位 / the linear location on an ascending axis
    IF fZ >= afZ[k] THEN // 已过该下节点 / the input is past this lower node
        nIz := k; // 记录候选单元 / register the candidate cell
    END_IF
END_FOR

// 段 5｜单元内归一化位置（单元宽度已证 > 0：轴严格升序 + 容差闸）/ segment 5, the normalised positions with a proven positive span
fX0 := afX[nIx]; // X 下节点 / the X lower node
fY0 := afY[nIy]; // Y 下节点 / the Y lower node
fZ0 := afZ[nIz]; // Z 下节点 / the Z lower node
fSpan := afX[nIx + 1] - fX0; // X 单元宽度 [用户单位] / the X cell span
IF fSpan <= DL_I3D_TOL THEN // 宽度非正（升序已证，属结构性不可达兜底）/ a non positive span, kept as a guard
    eErr := 16#0001_0627; // 故障级：轴向量退化，拒绝相除 / fault grade, the degenerate axis refuses the division
    bError := TRUE; // 置错误标志（R45 配对）/ raise the error flag, paired with the fault code
    bValid := FALSE; // 结果不可用 / the result void
    RETURN; // 早退 / early return
END_IF
fTx := (fX - fX0) / fSpan; // X 归一化位置（除子已证 > 容差）/ the X position with a proven divisor
fSpan := afY[nIy + 1] - fY0; // Y 单元宽度 [用户单位] / the Y cell span
IF fSpan <= DL_I3D_TOL THEN // 兜底闸 / the guard
    eErr := 16#0001_0627; // 故障级：轴向量退化 / fault grade, the degenerate axis
    bError := TRUE; // 置错误标志 / raise the error flag
    bValid := FALSE; // 结果不可用 / the result void
    RETURN; // 早退 / early return
END_IF
fTy := (fY - fY0) / fSpan; // Y 归一化位置 / the Y position
fSpan := afZ[nIz + 1] - fZ0; // Z 单元宽度 [用户单位] / the Z cell span
IF fSpan <= DL_I3D_TOL THEN // 兜底闸 / the guard
    eErr := 16#0001_0627; // 故障级：轴向量退化 / fault grade, the degenerate axis
    bError := TRUE; // 置错误标志 / raise the error flag
    bValid := FALSE; // 结果不可用 / the result void
    RETURN; // 早退 / early return
END_IF
fTz := (fZ - fZ0) / fSpan; // Z 归一化位置 / the Z position

// 段 6｜八角点取值与表值有限性（逐角点判，R272 数组侧覆盖）/ segment 6, the eight corners and the table finiteness
fC000 := afTable[nIx, nIy, nIz]; // 角点 000 / the corner 000
fC100 := afTable[nIx + 1, nIy, nIz]; // 角点 100 / the corner 100
fC010 := afTable[nIx, nIy + 1, nIz]; // 角点 010 / the corner 010
fC110 := afTable[nIx + 1, nIy + 1, nIz]; // 角点 110 / the corner 110
fC001 := afTable[nIx, nIy, nIz + 1]; // 角点 001 / the corner 001
fC101 := afTable[nIx + 1, nIy, nIz + 1]; // 角点 101 / the corner 101
fC011 := afTable[nIx, nIy + 1, nIz + 1]; // 角点 011 / the corner 011
fC111 := afTable[nIx + 1, nIy + 1, nIz + 1]; // 角点 111 / the corner 111
// 八角点逐个非有限判（覆盖本次参与的全部表值元素）/ the corner-wise non finite test over every participating value
IF (fC000 <> fC000) OR ((fC000 - fC000) <> (fC000 - fC000)) THEN // 角点 000 非有限 / the corner 000 is not finite
    bNonFin := TRUE; // 置非有限标记 / raise the non finite flag
END_IF
IF (fC100 <> fC100) OR ((fC100 - fC100) <> (fC100 - fC100)) THEN // 角点 100 非有限 / the corner 100 is not finite
    bNonFin := TRUE; // 置非有限标记 / raise the non finite flag
END_IF
IF (fC010 <> fC010) OR ((fC010 - fC010) <> (fC010 - fC010)) THEN // 角点 010 非有限 / the corner 010 is not finite
    bNonFin := TRUE; // 置非有限标记 / raise the non finite flag
END_IF
IF (fC110 <> fC110) OR ((fC110 - fC110) <> (fC110 - fC110)) THEN // 角点 110 非有限 / the corner 110 is not finite
    bNonFin := TRUE; // 置非有限标记 / raise the non finite flag
END_IF
IF (fC001 <> fC001) OR ((fC001 - fC001) <> (fC001 - fC001)) THEN // 角点 001 非有限 / the corner 001 is not finite
    bNonFin := TRUE; // 置非有限标记 / raise the non finite flag
END_IF
IF (fC101 <> fC101) OR ((fC101 - fC101) <> (fC101 - fC101)) THEN // 角点 101 非有限 / the corner 101 is not finite
    bNonFin := TRUE; // 置非有限标记 / raise the non finite flag
END_IF
IF (fC011 <> fC011) OR ((fC011 - fC011) <> (fC011 - fC011)) THEN // 角点 011 非有限 / the corner 011 is not finite
    bNonFin := TRUE; // 置非有限标记 / raise the non finite flag
END_IF
IF (fC111 <> fC111) OR ((fC111 - fC111) <> (fC111 - fC111)) THEN // 角点 111 非有限 / the corner 111 is not finite
    bNonFin := TRUE; // 置非有限标记 / raise the non finite flag
END_IF
IF bNonFin THEN // 表值含非有限 / a non finite table value exists
    eErr := 16#0001_0629; // 故障级：轴或表值含非有限值 / fault grade, a non finite axis or table value
    bError := TRUE; // 置错误标志（R45 配对）/ raise the error flag, paired with the fault code
    bValid := FALSE; // 结果不可用 / the result void
    FC_DL_InterpolateTable3D := 0.0; // 返回值回安全值 / the return back to the safe zero
    RETURN; // 早退 / early return
END_IF

// 段 7｜三线性插值 X→Y→Z（先沿最内维、再逐层，次序写死）/ segment 7, the trilinear interpolation with the fixed order
fA0 := fC000 + (fC100 - fC000) * fTx; // k 层 X 向插值 / the X interpolation on the lower layer
fA1 := fC001 + (fC101 - fC001) * fTx; // k+1 层 X 向插值 / the X interpolation on the upper layer
fB0 := fA0 + ((fC010 + (fC110 - fC010) * fTx) - fA0) * fTy; // k 层 Y 向插值 / the Y interpolation on the lower layer
fB1 := fA1 + ((fC011 + (fC111 - fC011) * fTx) - fA1) * fTy; // k+1 层 Y 向插值 / the Y interpolation on the upper layer
FC_DL_InterpolateTable3D := fB0 + (fB1 - fB0) * fTz; // Z 向插值出结果 / the Z interpolation gives the result

// 段 8｜结果复检兜底（非有限同拍三件套，边界四）/ segment 8, the result recheck with the triple on a non finite value
IF (FC_DL_InterpolateTable3D <> FC_DL_InterpolateTable3D)
OR ((FC_DL_InterpolateTable3D - FC_DL_InterpolateTable3D) <> (FC_DL_InterpolateTable3D - FC_DL_InterpolateTable3D)) THEN // 结果非有限 / the result is not finite
    FC_DL_InterpolateTable3D := 0.0; // 兜底安全值 / the bottom-line safe value
    eErr := 16#0001_0630; // 故障级：结果非有限（D9 返修独立码，不复用 0629）/ fault grade, the non finite result with its own code
    bError := TRUE; // 置错误标志（R45 配对）/ raise the error flag, paired with the fault code
    bValid := FALSE; // 结果不可用 / the result void
ELSE // 结果有限 / a finite result
    bValid := TRUE; // 结果可用 / the result is usable
END_IF
END_FUNCTION

(* ---- FC_DL_InterpStepNearest.st ---- *)
(*
    FC_DL_InterpStepNearest —— 查表最近邻（阶梯保持）插值（越界钳端点 + 并列取左邻）
    ------------------------------------------------------------------
    分类      : DL_MathData / Math-Interpolation
    前缀      : FC_DL_
    版本      : 1.0.0
    来源标签  : iec-std-wrapper（T0）
    溯源      : IEC 61131-3 标准语义的道莅防御性实现
                （纯查表比较逻辑，无内建插值内核依赖；未复制任何闭源厂商源码）
    平台      : 纯 IEC 61131-3，CODESYS / TwinCAT / InoProShop 通用
    分工声明  : 与存量 FC_DL_HermiteInterp / FC_DL_CubicSplineInterp /
                FC_DL_LagrangeInterp / FC_DL_InterpolateTable2D 分工——那四件
                为连续光滑或线性口径，本件为离散阶梯保持口径（最近邻，取整
                不平滑），越界端点钳位不外插。
    作者      : 道莅代码库 · PLC 编程专家（R57）
    ------------------------------------------------------------------
    功能说明  : 在按 x 升序排布的 n 点表中取最近邻 y（阶梯保持）。n 点 ≥2
                否则拒算；x 越界钳端点不外插；相邻 x 相等（表非单调）取先见
                点并置告警；距离并列取左邻（严格 < 判据，正中不摇摆）；
                非有限表项跳过并计数。
    错误码    : 0000 正常 / 16#0003_0007 点数不足拒算 / 16#0003_0008 表非单调告警 / 16#0003_0009 已钳端点
    修订记录  : 2026-11-21 v1.0.0 首次入库（R57 批 3 · 序号 15）
*)
FUNCTION FC_DL_InterpStepNearest : LREAL
VAR_IN_OUT
    afX : ARRAY[0..63] OF LREAL; // 表自变量数组 [工程单位]，升序排布 / the abscissa array, ascending
    afY : ARRAY[0..63] OF LREAL; // 表因变量数组 [工程单位] / the ordinate array
END_VAR
VAR_INPUT
    nCount  : DINT; // 表点数 [个]，域 2..64 / the point count, two through sixty four
    fXQuery : LREAL; // 查询自变量 [工程单位] / the query abscissa [engineering unit]
END_VAR
VAR_OUTPUT
    eErr    : UDINT; // 错误码，0 = 正常 / error code, zero is ok
    bError  : BOOL;  // 出错标志，eErr 非 0 时为真 / error flag, true when eErr is nonzero
    bValid  : BOOL;  // 结果是否为真实值，钳位/告警降级时为假 / the result is the true value, false when degraded
    bClamp  : BOOL;  // 发生端点钳位（不外插）[-] / an endpoint clamp happened, no extrapolation
    nSkipCnt: UDINT; // 跳过的非有限表项数 [个] / the skipped non finite table entries
END_VAR
VAR
    nI     : DINT;  // 循环计数 [个] / the loop counter
    nBest  : DINT;  // 最近点索引 [个] / the nearest index
    lrD    : LREAL; // 当前距离 [工程单位] / the current distance
    lrDbest: LREAL; // 当前最近距离 [工程单位] / the best distance so far
END_VAR

// 段 1｜返回值与错误状态预置安全值（四段式第一段，R45）/ segment 1, preset the return and error states
FC_DL_InterpStepNearest := 0.0; // 返回值预置安全值 0.0 / preset the return to the safe zero
eErr   := 16#0000_0000; // 错误码预置正常 / preset the code to ok
bError := FALSE; // 错误标志预置假 / preset the error flag false
bValid := TRUE; // 有效标志预置真 / preset the valid flag true
bClamp := FALSE; // 钳位标志预置假 / preset the clamp flag false
nSkipCnt := 0; // 跳过计数预置零 / preset the skip count zero

// 段 2｜点数域闸：n < 2 拒算（边界十五）/ segment 2, the count gate, below two rejects
IF nCount < 2 THEN // 点数不足 / insufficient points
    eErr   := 16#0003_0007; // 错误级：点数不足拒算 / error grade, insufficient points rejected
    bError := TRUE; // 置错误标志 / raise the error flag
    bValid := FALSE; // 输出不可用 / the output void
    RETURN; // 返回预置安全值 0.0 / return the preset safe zero
ELSIF nCount > 64 THEN // 超数组容量 / beyond the array capacity
    nCount := 64; // 钳到容量上限 / clamp to the capacity
    eErr   := 16#0003_0003; // 信息级：点数已钳位 / informational, the count clamped
    bError := TRUE; // 置错误标志 / raise the error flag
    bValid := FALSE; // 钳位口径非原始口径 / the clamped window is not the requested one
END_IF

// 段 3｜越界钳端点不外插（边界十五）/ segment 3, the endpoint clamp, no extrapolation
IF (fXQuery = fXQuery) AND ((fXQuery - fXQuery) = (fXQuery - fXQuery)) THEN // 查询值有限才判越界 / the clamp verdict only on a finite query
    IF fXQuery <= afX[0] THEN // 低于表首 / below the table head
        FC_DL_InterpStepNearest := afY[0]; // 钳端点返回 / clamp to the endpoint
        IF fXQuery < afX[0] THEN // 严格越界才置码 / the code only on a strict violation
            eErr   := 16#0003_0009; // 信息级：已钳下端点 / informational, clamped to the lower endpoint
            bError := TRUE; // 置错误标志 / raise the error flag
            bValid := FALSE; // 钳位结果非真实值 / the clamped result is not the true value
            bClamp := TRUE; // 置钳位标志 / raise the clamp flag
        END_IF
        RETURN; // 早退 / early return
    ELSIF fXQuery >= afX[nCount - 1] THEN // 高于表尾 / beyond the table tail
        FC_DL_InterpStepNearest := afY[nCount - 1]; // 钳端点返回 / clamp to the endpoint
        IF fXQuery > afX[nCount - 1] THEN // 严格越界才置码 / the code only on a strict violation
            eErr   := 16#0003_0009; // 信息级：已钳上端点 / informational, clamped to the upper endpoint
            bError := TRUE; // 置错误标志 / raise the error flag
            bValid := FALSE; // 钳位结果非真实值 / the clamped result is not the true value
            bClamp := TRUE; // 置钳位标志 / raise the clamp flag
        END_IF
        RETURN; // 早退 / early return
    END_IF
END_IF

// 段 4｜最近邻扫描：距离并列取左邻（严格 < 判据）/ segment 4, the nearest scan, ties take the left neighbor
nBest := 0; // 最近索引预置 0 / preset the nearest index
lrDbest := 1.7976931348623157E308; // 最近距离预置 LREAL 上界 / preset the best distance to the representable bound
FOR nI := 0 TO nCount - 1 DO // 有界循环 / the bounded loop
    IF (afX[nI] = afX[nI]) AND ((afX[nI] - afX[nI]) = (afX[nI] - afX[nI])) AND (afY[nI] = afY[nI]) AND ((afY[nI] - afY[nI]) = (afY[nI] - afY[nI])) THEN // 表项有限才参与 / only finite entries participate
        lrD := ABS(fXQuery - afX[nI]); // 当前距离 / the current distance
        IF lrD < lrDbest THEN // 严格小于才替换（并列保持左邻，正中不摇摆）/ strictly smaller replaces, ties hold the left
            lrDbest := lrD; // 更新最近距离 / update the best distance
            nBest := nI; // 更新最近索引 / update the nearest index
        END_IF
    ELSE // 非有限表项跳过 / a non finite entry skipped
        nSkipCnt := nSkipCnt + 1; // 跳过计数推进 / advance the skip count
    END_IF
END_FOR

// 段 5｜非单调告警与结果出口 / segment 5, the non monotonic warning and the outlet
FOR nI := 1 TO nCount - 1 DO // 相邻对扫查 / the adjacent pair scan
    IF (afX[nI] = afX[nI]) AND ((afX[nI] - afX[nI]) = (afX[nI] - afX[nI])) THEN // 有限项才比较 / finite entries only
        IF afX[nI] <= afX[nI - 1] THEN // 非递增即非单调 / a non increasing pair is non monotonic
            eErr   := 16#0003_0008; // 告警级：表非单调（先见点已按左邻规则保持）/ warning, a non monotonic table, the first seen held by the left rule
            bError := TRUE; // 置错误标志 / raise the error flag
            EXIT; // 一次告警即出 / one warning is enough
        END_IF
    END_IF
END_FOR
FC_DL_InterpStepNearest := afY[nBest]; // 最近邻 y 出口（阶梯保持）/ the nearest ordinate, the step hold
END_FUNCTION

(* ---- FC_DL_IntFloorLog2Udint.st ---- *)
(*==============================================================================
 * 组件名称 : FC_DL_IntFloorLog2Udint ｜ 子库 : DL_MathData ｜ v1.0.0 ｜ 2026-11-24
 * 平台     : CODESYS 3.5 / TwinCAT 3 / InoProShop / Machine Expert（纯 IEC，无厂商库）
 * 功能简介 : UDINT 下取整二进制对数 ⌊log2 nVal⌋。供位宽探测、二叉树层数、分频档位、
 *            哈希桶数 2 的幂归整使用。纯移位实现（逐次除 2 计数），禁浮点 LN，无精度问题。
 * 契约     : nVal ≥ 1 → 返回 0..31、bValid := TRUE；nVal = 0 → 返回 −1 且 bError := TRUE
 *            （log 在 0 处无定义，−1 为哨兵值而非合法结果，调用方必须查 bError）。
 * 依赖     : 无 DL_ 内部依赖（R16 自足实现），无标准库函数调用
 * 错误码   : R297 零码位范式：eErr 恒 0，仅以 bError / bValid 表达
 * 红线自检 : R1 零全局 R2 零%I/%Q R3 纯IEC R4 除零前置（被除数恒 2，无需域闸）+ 无浮点
 *            R5 双语注释 R6 N/A（无状态机）R7 N/A（无定时器/沿实例）
 *            R10 无类型转换 R11 全声明行分号 R15 标识符零保留字冲突
 * 遗留假设 : 返回值 −1 是故障哨兵，与「0 哨兵」范式不同：log2 的合法值含 0（nVal = 1），
 *            故不能用 0 表达故障；循环天然终止（nW 单调减半，最多 31 步），不设守卫。
 * 修订历史 : 2026-11-24 R79-B 首版（整数数论族补位）
 *============================================================================*)
FUNCTION FC_DL_IntFloorLog2Udint : DINT
VAR_INPUT
    nVal : UDINT := 0; // 待求对数的正整数 [无量纲] / the positive value whose binary logarithm is wanted
END_VAR
VAR_OUTPUT
    eErr   : UDINT; // 错误码，零码位范式恒 0 / error id, always zero under the zero-code rule
    bError : BOOL;  // 入参为零时为真 / TRUE when the argument is zero
    bValid : BOOL;  // 返回值可用标志 / TRUE when the return value is usable
END_VAR
VAR CONSTANT
    DL_ZERO : UDINT := 0; // 无符号零哨兵 / unsigned zero sentinel
    DL_ONE  : UDINT := 1; // 无符号一哨兵，循环终止阈值 / unsigned one, the loop exit threshold
    DL_TWO  : UDINT := 2; // 无符号二哨兵，移位基数 / unsigned two, the halving base
    DL_SENT : DINT  := -1; // 零入参故障哨兵 [无量纲] / the fault sentinel returned for a zero argument
    DL_ONEI : DINT  := 1;  // 整型一，计数步长 [次] / integer one, the counting step
    DL_NONE : DINT  := 0;  // 整型零，计数初值 [次] / integer zero, the counting start value
END_VAR
VAR
    nW   : UDINT; // 逐次减半的工作副本 [无量纲] / the working copy halved each pass
    nRes : DINT;  // 已减半次数，即 ⌊log2 nVal⌋ [次] / the number of halvings, that is the floor logarithm
END_VAR

// 段 1｜出口预置 / segment 1, preset the exit
FC_DL_IntFloorLog2Udint := DL_NONE;  // 缺省零 / default zero
eErr   := 0;                         // 零码位范式 / zero-code rule
bError := FALSE;                     // 预置无故障 / preset no fault
bValid := FALSE;                     // 域闸前不认返回值 / the return value is unusable until the gates pass

// 段 2｜零入参域闸：log2(0) 无定义，返回 −1 哨兵 / segment 2, the zero argument gate
IF nVal = DL_ZERO THEN
    FC_DL_IntFloorLog2Udint := DL_SENT;  // 故障哨兵 −1 / the fault sentinel minus one
    bError := TRUE;                      // 故障级 / fault level
    RETURN;                              // bValid 保持 FALSE / bValid stays FALSE
END_IF

// 段 3｜移位计数：nW 单调减半，nVal = 1 时零步即得 0 / segment 3, the halving count
nW   := nVal;                        // 工作副本 / the working copy
nRes := DL_NONE;                     // 计数清零 / clear the counter
WHILE nW > DL_ONE DO                 // 除零不可达：被除数恒为 2 / the divisor is the constant two
    nW   := nW / DL_TWO;             // 减半 / halve
    nRes := nRes + DL_ONEI;          // 计一次 / count one halving
END_WHILE

// 段 4｜出口 / segment 4, the exit
FC_DL_IntFloorLog2Udint := nRes;     // 回写 ⌊log2 nVal⌋ / publish the floor logarithm
bValid := TRUE;                      // 返回值可用 / the return value is usable
END_FUNCTION

(* ---- FC_DL_IntIsPerfectSquareUdint.st ---- *)
(*==============================================================================
 * 组件名称 : FC_DL_IntIsPerfectSquareUdint ｜ 子库 : DL_MathData ｜ v1.0.0 ｜ 2026-11-24
 * 平台     : CODESYS 3.5 / TwinCAT 3 / InoProShop / Machine Expert（纯 IEC，无厂商库）
 * 功能简介 : 判定无符号整数是否为完全平方数。先牛顿迭代求 ⌊√nVal⌋，再回乘比较 ——
 *            回乘前先判根是否 > 65535：UDINT 域内平方根最大 65535，越界者
 *            平方必超 2^32，回乘会回绕，故直接判否（溢出结构性拦在乘法之前）。
 * 契约     : 返回 TRUE=完全平方数（0 视为完全平方）；迭代未收敛时置 bError 并返回 FALSE。
 * 依赖     : 无 DL_ 内部依赖（R16 自足实现），无标准库函数调用
 * 错误码   : R297 零码位范式：eErr 恒 0，仅以 bError / bValid 表达
 * 红线自检 : R1 零全局 R2 零%I/%Q R3 纯IEC R4 回乘前溢出反算 + 迭代上限 + 除零前置
 *            R5 双语注释 R6 N/A（无状态机）R7 N/A（无定时器/沿实例）
 *            R10 无类型转换 R11 全声明行分号 R15 标识符零保留字冲突 R18 N/A（无 bReset）
 * 修订历史 : 2026-11-24 R79-A 首版（整数数论族 2/8）
 *============================================================================*)
FUNCTION FC_DL_IntIsPerfectSquareUdint : BOOL
VAR_INPUT
    nVal        : UDINT;    // 待判定整数，全域 0~16#FFFF_FFFF [无量纲] / candidate over the whole unsigned range
END_VAR
VAR_OUTPUT
    eErr        : UDINT;    // 错误码，零码位范式恒 0 / error id, always zero under the zero-code rule
    bError      : BOOL;     // 迭代未收敛为真（结构性不可达） / TRUE when the iteration fails to converge, unreachable in theory
    bValid      : BOOL;     // 判定可用标志 / TRUE when the verdict is usable
END_VAR
VAR CONSTANT
    DL_TWO      : UDINT := 2;               // 牛顿迭代除数 [无量纲] / Newton divisor, dimensionless
    DL_ONE      : UDINT := 1;               // 整数一 [无量纲] / integer one, dimensionless
    DL_ZERO     : UDINT := 0;               // 整数零哨兵 [无量纲] / integer zero sentinel, dimensionless
    DL_ITER_MAX : UDINT := 64;              // 迭代次数上限 [次] / iteration cap [count]
    DL_ROOT_MAX : UDINT := 65535;           // UDINT 域内平方根上限，超过则平方必溢出 [无量纲] / largest root that still squares inside the unsigned range
END_VAR
VAR
    nApprox     : UDINT;    // 当前试值 / current trial value
    nNext       : UDINT;    // 下一试值 / next trial value
    nIter       : UDINT;    // 已用迭代次数 / iterations consumed so far
    nSquare     : UDINT;    // 根的回乘结果 / square of the resolved root
END_VAR

// 段 1｜出口预置 / segment 1, preset the exit
FC_DL_IntIsPerfectSquareUdint := FALSE;     // 缺省非完全平方 / default not a perfect square
eErr   := 0;                                // 零码位范式 / zero-code rule
bError := FALSE;                            // 预置无故障 / preset no fault
bValid := FALSE;                            // 迭代结束前不认判定 / unusable until the iteration ends

// 段 2｜零边界：0 = 0²，直接判真 / segment 2, the zero boundary
IF nVal = DL_ZERO THEN
    bValid := TRUE;                         // 判定可用 / the verdict is usable
    FC_DL_IntIsPerfectSquareUdint := TRUE;  // 零是完全平方 / zero is a perfect square
    RETURN;
END_IF

// 段 3｜牛顿迭代求根（与求根族同法，内联自足不跨件调用） / segment 3, inline Newton root
nApprox := (nVal / DL_TWO) + DL_ONE;        // 上界初值 / upper bound start
nIter   := DL_ZERO;
WHILE nIter < DL_ITER_MAX DO
    nIter := nIter + DL_ONE;                // 计数 / count
    nNext := (nApprox + (nVal / nApprox)) / DL_TWO;    // 下一试值 / next trial
    IF nNext >= nApprox THEN
        EXIT;                               // 收敛 / converged
    END_IF
    nApprox := nNext;
END_WHILE
IF nIter >= DL_ITER_MAX THEN
    bError := TRUE;                         // 未收敛（理论不可达）/ not converged, unreachable in theory
    RETURN;                                 // 返回 FALSE 且 bValid 保持 FALSE / return FALSE with bValid still FALSE
END_IF

// 段 4｜回乘比较：先拦溢出再乘 / segment 4, overflow reflection before the multiplication
IF nApprox > DL_ROOT_MAX THEN
    bValid := TRUE;                         // 判定成立：根超 65535 必非域内平方 / a root above 65535 cannot square inside the domain
    RETURN;                                 // 返回 FALSE / return FALSE
END_IF
nSquare := nApprox * nApprox;               // 根 ≤ 65535，平方 ≤ 16#FFFE_0001 不溢出 / the square stays inside the unsigned range
IF nSquare = nVal THEN
    FC_DL_IntIsPerfectSquareUdint := TRUE;  // 回乘相等即完全平方 / an equal square proves the verdict
END_IF
bValid := TRUE;                             // 判定可用 / the verdict is usable
END_FUNCTION
